(* IEC 61131-3 sources: plc-st-coding-agent/progress/evidence/f14_v10_full_20261113/jobs/custom_minimax-m27 (part 5) *)

(* ---- public-medium-05.candidate_02.st ---- *)
(* ENGINEERING_CONTRACT *)
(*
  PubRefs: PUB001, PUB003, PUB004, PUB006, PUB007
  Mode: 0=manual, 1=automatic
  Manual (Mode=FALSE): ForwardButton→MotorForward, ReverseButton→MotorReverse; interlocked (PUB001)
  Auto (Mode=TRUE):
    IDLE+SensorA→WAIT_AT_A (PUB003)
    WAIT_AT_A+ButtonA→MOVING_AB; MotorForward=TRUE (PUB003)
    MOVING_AB+SensorB→WAIT_AT_B; MotorForward=FALSE (PUB004)
    WAIT_AT_B+ButtonB→MOVING_BC; MotorForward=TRUE (PUB004)
    MOVING_BC+SensorC→WAIT_AT_C; MotorForward=FALSE (PUB004)
    WAIT_AT_C+ButtonC→COMPLETE; CompletionLight=TRUE (PUB006)
    COMPLETE+NOT SensorC→IDLE; CompletionLight=FALSE (PUB007)
  Retention: CompletionLight holds until SensorC clears (PUB007)
  Reset on mode switch: Auto state→IDLE, motor OFF
*)
(* CONTRACT_RULES [] *)

TYPE ProdState :
(
    IDLE      := 0,
    WAIT_AT_A := 1,
    MOVING_AB := 2,
    WAIT_AT_B := 3,
    MOVING_BC := 4,
    WAIT_AT_C := 5,
    COMPLETE  := 6
);
END_TYPE;

FUNCTION_BLOCK ProdLineControl
VAR_INPUT
    Mode          : BOOL;
    ForwardButton : BOOL;
    ReverseButton : BOOL;
    SensorA       : BOOL;
    SensorB       : BOOL;
    SensorC       : BOOL;
    ButtonA       : BOOL;
    ButtonB       : BOOL;
    ButtonC       : BOOL;
END_VAR
VAR
    tmp_State : ProdState := IDLE;
END_VAR
VAR_OUTPUT
    MotorForward    : BOOL := FALSE;
    MotorReverse    : BOOL := FALSE;
    CompletionLight : BOOL := FALSE;
END_VAR

// --- Automatic Mode State Machine ---
IF Mode THEN
    CASE tmp_State OF
        IDLE :
            MotorForward    := FALSE;
            MotorReverse    := FALSE;
            CompletionLight := FALSE;
            IF SensorA THEN
                tmp_State := WAIT_AT_A;
            END_IF;

        WAIT_AT_A :
            MotorForward    := FALSE;
            MotorReverse    := FALSE;
            CompletionLight := FALSE;
            IF ButtonA THEN
                tmp_State := MOVING_AB;
            END_IF;

        MOVING_AB :
            MotorForward    := TRUE;
            MotorReverse    := FALSE;
            CompletionLight := FALSE;
            IF SensorB THEN
                tmp_State     := WAIT_AT_B;
                MotorForward  := FALSE;
            END_IF;

        WAIT_AT_B :
            MotorForward    := FALSE;
            MotorReverse    := FALSE;
            CompletionLight := FALSE;
            IF ButtonB THEN
                tmp_State := MOVING_BC;
            END_IF;

        MOVING_BC :
            MotorForward    := TRUE;
            MotorReverse    := FALSE;
            CompletionLight := FALSE;
            IF SensorC THEN
                tmp_State     := WAIT_AT_C;
                MotorForward  := FALSE;
            END_IF;

        WAIT_AT_C :
            MotorForward    := FALSE;
            MotorReverse    := FALSE;
            IF ButtonC THEN
                tmp_State       := COMPLETE;
                CompletionLight := TRUE;
            END_IF;

        COMPLETE :
            MotorForward    := FALSE;
            MotorReverse    := FALSE;
            CompletionLight := TRUE;
            IF NOT SensorC THEN
                tmp_State       := IDLE;
                CompletionLight := FALSE;
            END_IF;
    END_CASE;

// --- Manual Mode ---
ELSE
    MotorForward := ForwardButton AND NOT ReverseButton;
    MotorReverse := ReverseButton AND NOT ForwardButton;
    tmp_State    := IDLE;
END_IF;

END_FUNCTION_BLOCK

(* ---- public-medium-05.raw_candidate_01.st ---- *)
(* ENGINEERING_CONTRACT *)
(*
  PubRefs: PUB001, PUB003, PUB004, PUB006, PUB007
  Mode: 0=manual, 1=automatic
  Manual (Mode=FALSE): ForwardButton→MotorForward, ReverseButton→MotorReverse; interlocked (PUB001)
  Auto (Mode=TRUE):
    IDLE+SensorA→WAIT_AT_A (PUB003)
    WAIT_AT_A+ButtonA→MOVING_AB; MotorForward=TRUE (PUB003)
    MOVING_AB+SensorB→WAIT_AT_B; MotorForward=FALSE (PUB004)
    WAIT_AT_B+ButtonB→MOVING_BC; MotorForward=TRUE (PUB004)
    MOVING_BC+SensorC→WAIT_AT_C; MotorForward=FALSE (PUB004)
    WAIT_AT_C+ButtonC→COMPLETE; CompletionLight=TRUE (PUB006)
    COMPLETE+NOT SensorC→IDLE; CompletionLight=FALSE (PUB007)
  Retention: CompletionLight holds until SensorC clears (PUB007)
  Reset on mode switch: Auto state→IDLE, motor OFF
*)
(* CONTRACT_RULES [] *)

TYPE ProdState :
(
    IDLE      := 0,
    WAIT_AT_A := 1,
    MOVING_AB := 2,
    WAIT_AT_B := 3,
    MOVING_BC := 4,
    WAIT_AT_C := 5,
    COMPLETE  := 6
);
END_TYPE

FUNCTION_BLOCK ProdLineControl
VAR
    tmp_State : ProdState := IDLE;
END_VAR
VAR_OUTPUT
    MotorForward    : BOOL := FALSE;
    MotorReverse    : BOOL := FALSE;
    CompletionLight : BOOL := FALSE;
END_VAR

// --- Automatic Mode State Machine ---
IF Mode THEN
    CASE tmp_State OF
        IDLE :
            MotorForward    := FALSE;
            MotorReverse    := FALSE;
            CompletionLight := FALSE;
            IF SensorA THEN
                tmp_State := WAIT_AT_A;
            END_IF;

        WAIT_AT_A :
            MotorForward    := FALSE;
            MotorReverse    := FALSE;
            CompletionLight := FALSE;
            IF ButtonA THEN
                tmp_State := MOVING_AB;
            END_IF;

        MOVING_AB :
            MotorForward    := TRUE;
            MotorReverse    := FALSE;
            CompletionLight := FALSE;
            IF SensorB THEN
                tmp_State     := WAIT_AT_B;
                MotorForward  := FALSE;
            END_IF;

        WAIT_AT_B :
            MotorForward    := FALSE;
            MotorReverse    := FALSE;
            CompletionLight := FALSE;
            IF ButtonB THEN
                tmp_State := MOVING_BC;
            END_IF;

        MOVING_BC :
            MotorForward    := TRUE;
            MotorReverse    := FALSE;
            CompletionLight := FALSE;
            IF SensorC THEN
                tmp_State     := WAIT_AT_C;
                MotorForward  := FALSE;
            END_IF;

        WAIT_AT_C :
            MotorForward    := FALSE;
            MotorReverse    := FALSE;
            IF ButtonC THEN
                tmp_State      := COMPLETE;
                CompletionLight := TRUE;
            END_IF;

        COMPLETE :
            MotorForward    := FALSE;
            MotorReverse    := FALSE;
            CompletionLight := TRUE;
            IF NOT SensorC THEN
                tmp_State      := IDLE;
                CompletionLight := FALSE;
            END_IF;
    END_CASE;

// --- Manual Mode ---
ELSE
    MotorForward := ForwardButton AND NOT ReverseButton;
    MotorReverse := ReverseButton AND NOT ForwardButton;
    tmp_State    := IDLE;
END_IF;

END_FUNCTION_BLOCK

(* ---- public-medium-05.raw_candidate_02.st ---- *)
(* ENGINEERING_CONTRACT *)
(*
  PubRefs: PUB001, PUB003, PUB004, PUB006, PUB007
  Mode: 0=manual, 1=automatic
  Manual (Mode=FALSE): ForwardButton→MotorForward, ReverseButton→MotorReverse; interlocked (PUB001)
  Auto (Mode=TRUE):
    IDLE+SensorA→WAIT_AT_A (PUB003)
    WAIT_AT_A+ButtonA→MOVING_AB; MotorForward=TRUE (PUB003)
    MOVING_AB+SensorB→WAIT_AT_B; MotorForward=FALSE (PUB004)
    WAIT_AT_B+ButtonB→MOVING_BC; MotorForward=TRUE (PUB004)
    MOVING_BC+SensorC→WAIT_AT_C; MotorForward=FALSE (PUB004)
    WAIT_AT_C+ButtonC→COMPLETE; CompletionLight=TRUE (PUB006)
    COMPLETE+NOT SensorC→IDLE; CompletionLight=FALSE (PUB007)
  Retention: CompletionLight holds until SensorC clears (PUB007)
  Reset on mode switch: Auto state→IDLE, motor OFF
*)
(* CONTRACT_RULES [] *)

TYPE ProdState :
(
    IDLE      := 0,
    WAIT_AT_A := 1,
    MOVING_AB := 2,
    WAIT_AT_B := 3,
    MOVING_BC := 4,
    WAIT_AT_C := 5,
    COMPLETE  := 6
);
END_TYPE;

FUNCTION_BLOCK ProdLineControl
VAR_INPUT
    Mode          : BOOL;
    ForwardButton : BOOL;
    ReverseButton : BOOL;
    SensorA       : BOOL;
    SensorB       : BOOL;
    SensorC       : BOOL;
    ButtonA       : BOOL;
    ButtonB       : BOOL;
    ButtonC       : BOOL;
END_VAR
VAR
    tmp_State : ProdState := IDLE;
END_VAR
VAR_OUTPUT
    MotorForward    : BOOL := FALSE;
    MotorReverse    : BOOL := FALSE;
    CompletionLight : BOOL := FALSE;
END_VAR

// --- Automatic Mode State Machine ---
IF Mode THEN
    CASE tmp_State OF
        IDLE :
            MotorForward    := FALSE;
            MotorReverse    := FALSE;
            CompletionLight := FALSE;
            IF SensorA THEN
                tmp_State := WAIT_AT_A;
            END_IF;

        WAIT_AT_A :
            MotorForward    := FALSE;
            MotorReverse    := FALSE;
            CompletionLight := FALSE;
            IF ButtonA THEN
                tmp_State := MOVING_AB;
            END_IF;

        MOVING_AB :
            MotorForward    := TRUE;
            MotorReverse    := FALSE;
            CompletionLight := FALSE;
            IF SensorB THEN
                tmp_State     := WAIT_AT_B;
                MotorForward  := FALSE;
            END_IF;

        WAIT_AT_B :
            MotorForward    := FALSE;
            MotorReverse    := FALSE;
            CompletionLight := FALSE;
            IF ButtonB THEN
                tmp_State := MOVING_BC;
            END_IF;

        MOVING_BC :
            MotorForward    := TRUE;
            MotorReverse    := FALSE;
            CompletionLight := FALSE;
            IF SensorC THEN
                tmp_State     := WAIT_AT_C;
                MotorForward  := FALSE;
            END_IF;

        WAIT_AT_C :
            MotorForward    := FALSE;
            MotorReverse    := FALSE;
            IF ButtonC THEN
                tmp_State       := COMPLETE;
                CompletionLight := TRUE;
            END_IF;

        COMPLETE :
            MotorForward    := FALSE;
            MotorReverse    := FALSE;
            CompletionLight := TRUE;
            IF NOT SensorC THEN
                tmp_State       := IDLE;
                CompletionLight := FALSE;
            END_IF;
    END_CASE;

// --- Manual Mode ---
ELSE
    MotorForward := ForwardButton AND NOT ReverseButton;
    MotorReverse := ReverseButton AND NOT ForwardButton;
    tmp_State    := IDLE;
END_IF;

END_FUNCTION_BLOCK

(* ---- public-medium-06.candidate_01.st ---- *)
(* ENGINEERING_CONTRACT *)
(*
| Output/State            | Activation              | Retention          | Reset/Deactivation                | Same-scan Priority | Units/Boundaries     |
|-------------------------|-------------------------|--------------------|-----------------------------------|--------------------|----------------------|
| THICKNESS_ALARM         | Immediate on valid TRUE | Hold >=500ms min   | Signal invalid OR hold timer done | Alarm active wins  | TON PT=500ms         |
| Slab_Fault_Counter      | Rising edge of valid    | Count accumulates  | Power-up only                     | N/A                | UINT max             |
| Slab_Fault_History[0]   | Rising edge of valid    | Newest entry       | Power-up only                     | N/A                | DINT timestamp       |
| Slab_Fault_History[1-4] | Shifted from lower idx  | Older entries      | Power-up only                     | N/A                | DINT timestamp       |
| Slab_Runtime_Accumulator| Accum when cutting valid| Accumulates       | Power-up only                     | N/A                | LTIME nanoseconds    |
| Hold timer (TON)        | Starts on fault clear   | Runs for PT        | Q=TRUE stops hold; signal invalid | N/A                | PT=T#500ms           |
| prev_valid_fault (VAR)  | Updated each scan       | Last cycle fault   | Power-up only                     | N/A                | BOOL                 |
| alarm_state (VAR)       | Transitions per FSM     | Holds across scans | Signal invalid resets             | N/A                | (0,1,2) enum         |
*)
(* CONTRACT_RULES [] *)

TYPE AlarmState :
(
    AlarmOff    := 0,
    FaultActive := 1,
    FaultCleared := 2
);
END_TYPE;

FUNCTION_BLOCK SlabThicknessMonitor
    VAR_INPUT
        THICKNESS_FAULT        : BOOL;
        THICKNESS_SIGNAL_VALID : BOOL;
        CUTTING_RUN            : BOOL;
        FaultTimestamp         : DINT;
        CycleTime              : TIME;
    END_VAR
    VAR_OUTPUT
        THICKNESS_ALARM         : BOOL := FALSE;
        Slab_Fault_Counter      : UINT := 0;
        Slab_Runtime_Accumulator: LTIME := LTIME#0s;
        Slab_Fault_History      : ARRAY[0..4] OF DINT := [5(DINT#0)];
    END_VAR
    VAR
        prev_valid_fault : BOOL := FALSE;
        hold_timer       : TON;
        alarm_state      : AlarmState := AlarmOff;
        tmp_hold_q       : BOOL;
    END_VAR

    // Clear all state when signal becomes invalid (power-up also covered by first-scan initialization)
    IF NOT THICKNESS_SIGNAL_VALID THEN
        alarm_state         := AlarmOff;
        THICKNESS_ALARM     := FALSE;
        hold_timer(IN := FALSE);
        prev_valid_fault    := FALSE;
        Slab_Fault_Counter  := 0;
        Slab_Fault_History  := [5(DINT#0)];
        Slab_Runtime_Accumulator := LTIME#0s;
    ELSE
        // Detect FALSE-to-TRUE transition of valid fault signal (PUB001)
        IF prev_valid_fault = FALSE AND THICKNESS_FAULT = TRUE THEN
            // Shift history: older entries toward higher indices, retain 5 most recent
            Slab_Fault_History[4] := Slab_Fault_History[3];
            Slab_Fault_History[3] := Slab_Fault_History[2];
            Slab_Fault_History[2] := Slab_Fault_History[1];
            Slab_Fault_History[1] := Slab_Fault_History[0];
            Slab_Fault_History[0] := FaultTimestamp;
            Slab_Fault_Counter := Slab_Fault_Counter + UINT#1;
        END_IF;

        // Accumulate runtime only while cutting, signal valid, no fault (PUB003)
        IF CUTTING_RUN AND NOT THICKNESS_FAULT THEN
            Slab_Runtime_Accumulator := Slab_Runtime_Accumulator + CycleTime;
        END_IF;

        // Alarm state machine with 500ms minimum hold (PUB001, PUB002)
        // Evaluate timer first so same-scan enable and elapsed origin agree
        hold_timer(IN := (alarm_state = FaultCleared));
        tmp_hold_q := hold_timer.Q;

        CASE alarm_state OF
            AlarmOff:
                IF THICKNESS_FAULT THEN
                    alarm_state     := FaultActive;
                    THICKNESS_ALARM := TRUE;
                END_IF;

            FaultActive:
                THICKNESS_ALARM := TRUE;
                IF NOT THICKNESS_FAULT THEN
                    alarm_state := FaultCleared;
                END_IF;

            FaultCleared:
                THICKNESS_ALARM := TRUE;
                IF tmp_hold_q THEN
                    alarm_state     := AlarmOff;
                    THICKNESS_ALARM := FALSE;
                END_IF;
        END_CASE;
    END_IF;

    // Update previous fault state for next scan edge detection
    prev_valid_fault := THICKNESS_FAULT;
END_FUNCTION_BLOCK

(* ---- public-medium-06.candidate_02.st ---- *)
(* ENGINEERING_CONTRACT *)
(*
| Output/State            | Activation              | Retention          | Reset/Deactivation                | Same-scan Priority | Units/Boundaries     |
|-------------------------|-------------------------|--------------------|-----------------------------------|--------------------|----------------------|
| THICKNESS_ALARM         | Immediate on valid TRUE | Hold >=500ms min   | Signal invalid OR hold timer done | Alarm active wins  | TON PT=500ms         |
| Slab_Fault_Counter      | Rising edge of valid    | Count accumulates  | Power-up only                     | N/A                | UINT max             |
| Slab_Fault_History[0]   | Rising edge of valid    | Newest entry       | Power-up only                     | N/A                | DINT timestamp       |
| Slab_Fault_History[1-4] | Shifted from lower idx  | Older entries      | Power-up only                     | N/A                | DINT timestamp       |
| Slab_Runtime_Accumulator| Accum when cutting valid| Accumulates       | Power-up only                     | N/A                | LTIME nanoseconds    |
| Hold timer (TON)        | Starts on fault clear   | Runs for PT        | Q=TRUE stops hold; signal invalid | N/A                | PT=T#500ms           |
| prev_valid_fault (VAR)  | Updated each scan       | Last cycle fault   | Power-up only                     | N/A                | BOOL                 |
| alarm_state (VAR)       | Transitions per FSM     | Holds across scans | Signal invalid resets             | N/A                | (0,1,2) enum         |
*)
(* CONTRACT_RULES [] *)

TYPE AlarmState :
(
    AlarmOff    := 0,
    FaultActive := 1,
    FaultCleared := 2
);
END_TYPE;

FUNCTION_BLOCK SlabThicknessMonitor
    VAR_INPUT
        THICKNESS_FAULT        : BOOL;
        THICKNESS_SIGNAL_VALID : BOOL;
        CUTTING_RUN            : BOOL;
        FaultTimestamp         : DINT;
        CycleTime              : TIME;
    END_VAR
    VAR_OUTPUT
        THICKNESS_ALARM         : BOOL := FALSE;
        Slab_Fault_Counter      : UINT := 0;
        Slab_Runtime_Accumulator: LTIME := LTIME#0s;
        Slab_Fault_History      : ARRAY[0..4] OF DINT := [DINT#0, DINT#0, DINT#0, DINT#0, DINT#0];
    END_VAR
    VAR
        prev_valid_fault : BOOL := FALSE;
        hold_timer       : TON;
        alarm_state      : AlarmState := AlarmOff;
        tmp_hold_q       : BOOL;
    END_VAR

    // Clear all state when signal becomes invalid (power-up also covered by first-scan initialization)
    IF NOT THICKNESS_SIGNAL_VALID THEN
        alarm_state         := AlarmOff;
        THICKNESS_ALARM     := FALSE;
        hold_timer(IN := FALSE);
        prev_valid_fault    := FALSE;
        Slab_Fault_Counter  := 0;
        Slab_Fault_History  := [DINT#0, DINT#0, DINT#0, DINT#0, DINT#0];
        Slab_Runtime_Accumulator := LTIME#0s;
    ELSE
        // Detect FALSE-to-TRUE transition of valid fault signal (PUB001)
        IF prev_valid_fault = FALSE AND THICKNESS_FAULT = TRUE THEN
            // Shift history: older entries toward higher indices, retain 5 most recent
            Slab_Fault_History[4] := Slab_Fault_History[3];
            Slab_Fault_History[3] := Slab_Fault_History[2];
            Slab_Fault_History[2] := Slab_Fault_History[1];
            Slab_Fault_History[1] := Slab_Fault_History[0];
            Slab_Fault_History[0] := FaultTimestamp;
            Slab_Fault_Counter := Slab_Fault_Counter + UINT#1;
        END_IF;

        // Accumulate runtime only while cutting, signal valid, no fault (PUB003)
        IF CUTTING_RUN AND NOT THICKNESS_FAULT THEN
            Slab_Runtime_Accumulator := Slab_Runtime_Accumulator + CycleTime;
        END_IF;

        // Alarm state machine with 500ms minimum hold (PUB001, PUB002)
        // Evaluate timer first so same-scan enable and elapsed origin agree
        hold_timer(IN := (alarm_state = FaultCleared));
        tmp_hold_q := hold_timer.Q;

        CASE alarm_state OF
            AlarmOff:
                IF THICKNESS_FAULT THEN
                    alarm_state     := FaultActive;
                    THICKNESS_ALARM := TRUE;
                END_IF;

            FaultActive:
                THICKNESS_ALARM := TRUE;
                IF NOT THICKNESS_FAULT THEN
                    alarm_state := FaultCleared;
                END_IF;

            FaultCleared:
                THICKNESS_ALARM := TRUE;
                IF tmp_hold_q THEN
                    alarm_state     := AlarmOff;
                    THICKNESS_ALARM := FALSE;
                END_IF;
        END_CASE;
    END_IF;

    // Update previous fault state for next scan edge detection
    prev_valid_fault := THICKNESS_FAULT;
END_FUNCTION_BLOCK

(* ---- public-medium-06.candidate_03.st ---- *)
(* ENGINEERING_CONTRACT *)
(*
| Output/State            | Activation              | Retention          | Reset/Deactivation                | Same-scan Priority | Units/Boundaries     |
|-------------------------|-------------------------|--------------------|-----------------------------------|--------------------|----------------------|
| THICKNESS_ALARM         | Immediate on valid TRUE | Hold >=500ms min   | Signal invalid OR hold timer done | Alarm active wins  | TON PT=500ms         |
| Slab_Fault_Counter      | Rising edge of valid    | Count accumulates  | Power-up only                     | N/A                | UINT max             |
| Slab_Fault_History[0]   | Rising edge of valid    | Newest entry       | Power-up only                     | N/A                | DINT timestamp       |
| Slab_Fault_History[1-4] | Shifted from lower idx  | Older entries      | Power-up only                     | N/A                | DINT timestamp       |
| Slab_Runtime_Accumulator| Accum when cutting valid| Accumulates       | Power-up only                     | N/A                | LTIME nanoseconds    |
| Hold timer (TON)        | Starts on fault clear   | Runs for PT        | Q=TRUE stops hold; signal invalid | N/A                | PT=T#500ms           |
| prev_valid_fault (VAR)  | Updated each scan       | Last cycle fault   | Power-up only                     | N/A                | BOOL                 |
| alarm_state (VAR)       | Transitions per FSM     | Holds across scans | Signal invalid resets             | N/A                | (0,1,2) enum         |
*)
(* CONTRACT_RULES [] *)

TYPE AlarmState :
(
    AlarmOff    := 0,
    FaultActive := 1,
    FaultCleared := 2
);
END_TYPE;

FUNCTION_BLOCK SlabThicknessMonitor
    VAR_INPUT
        THICKNESS_FAULT        : BOOL;
        THICKNESS_SIGNAL_VALID : BOOL;
        CUTTING_RUN            : BOOL;
        FaultTimestamp         : DINT;
        CycleTime              : TIME;
    END_VAR
    VAR_OUTPUT
        THICKNESS_ALARM         : BOOL := FALSE;
        Slab_Fault_Counter      : UINT := 0;
        Slab_Runtime_Accumulator: LTIME := LTIME#0s;
        Slab_Fault_History      : ARRAY[0..4] OF DINT;
    END_VAR
    VAR
        prev_valid_fault : BOOL := FALSE;
        hold_timer       : TON;
        alarm_state      : AlarmState := AlarmOff;
        tmp_hold_q       : BOOL;
        tmp_idx          : UINT;
    END_VAR

    // Clear all state when signal becomes invalid (power-up also covered by first-scan initialization)
    IF NOT THICKNESS_SIGNAL_VALID THEN
        alarm_state         := AlarmOff;
        THICKNESS_ALARM     := FALSE;
        hold_timer(IN := FALSE);
        prev_valid_fault    := FALSE;
        Slab_Fault_Counter  := 0;
        Slab_Fault_History[0] := DINT#0;
        Slab_Fault_History[1] := DINT#0;
        Slab_Fault_History[2] := DINT#0;
        Slab_Fault_History[3] := DINT#0;
        Slab_Fault_History[4] := DINT#0;
        Slab_Runtime_Accumulator := LTIME#0s;
    ELSE
        // Detect FALSE-to-TRUE transition of valid fault signal (PUB001)
        IF prev_valid_fault = FALSE AND THICKNESS_FAULT = TRUE THEN
            // Shift history: older entries toward higher indices, retain 5 most recent
            Slab_Fault_History[4] := Slab_Fault_History[3];
            Slab_Fault_History[3] := Slab_Fault_History[2];
            Slab_Fault_History[2] := Slab_Fault_History[1];
            Slab_Fault_History[1] := Slab_Fault_History[0];
            Slab_Fault_History[0] := FaultTimestamp;
            Slab_Fault_Counter := Slab_Fault_Counter + UINT#1;
        END_IF;

        // Accumulate runtime only while cutting, signal valid, no fault (PUB003)
        IF CUTTING_RUN AND NOT THICKNESS_FAULT THEN
            Slab_Runtime_Accumulator := Slab_Runtime_Accumulator + CycleTime;
        END_IF;

        // Alarm state machine with 500ms minimum hold (PUB001, PUB002)
        // Evaluate timer first so same-scan enable and elapsed origin agree
        hold_timer(IN := (alarm_state = FaultCleared));
        tmp_hold_q := hold_timer.Q;

        CASE alarm_state OF
            AlarmOff:
                IF THICKNESS_FAULT THEN
                    alarm_state     := FaultActive;
                    THICKNESS_ALARM := TRUE;
                END_IF;

            FaultActive:
                THICKNESS_ALARM := TRUE;
                IF NOT THICKNESS_FAULT THEN
                    alarm_state := FaultCleared;
                END_IF;

            FaultCleared:
                THICKNESS_ALARM := TRUE;
                IF tmp_hold_q THEN
                    alarm_state     := AlarmOff;
                    THICKNESS_ALARM := FALSE;
                END_IF;
        END_CASE;
    END_IF;

    // Update previous fault state for next scan edge detection
    prev_valid_fault := THICKNESS_FAULT;
END_FUNCTION_BLOCK

(* ---- public-medium-06.candidate_04.st ---- *)
(* ENGINEERING_CONTRACT *)
(*
| Output/State            | Activation              | Retention          | Reset/Deactivation                | Same-scan Priority | Units/Boundaries     |
|-------------------------|-------------------------|--------------------|-----------------------------------|--------------------|----------------------|
| THICKNESS_ALARM         | Immediate on valid TRUE | Hold >=500ms min   | Signal invalid OR hold timer done | Alarm active wins  | TON PT=T#500ms       |
| Slab_Fault_Counter      | Rising edge of valid    | Count accumulates  | Power-up only                     | N/A                | UINT max             |
| Slab_Fault_History[0]   | Rising edge of valid    | Newest entry       | Power-up only                     | N/A                | DINT timestamp       |
| Slab_Fault_History[1-4] | Shifted from lower idx  | Older entries      | Power-up only                     | N/A                | DINT timestamp       |
| Slab_Runtime_Accumulator| Accum when cutting valid| Accumulates       | Power-up only                     | N/A                | LTIME nanoseconds    |
| Hold timer (TON)        | Starts on fault clear   | Runs for PT        | Q=TRUE stops hold; signal invalid | N/A                | PT=T#500ms           |
| prev_valid_fault (VAR)  | Updated each scan       | Last cycle fault   | Power-up only                     | N/A                | BOOL                 |
| alarm_state (VAR)       | Transitions per FSM     | Holds across scans | Signal invalid resets             | N/A                | (0,1,2) enum         |
*)
(* CONTRACT_RULES [] *)

TYPE AlarmState :
(
    AlarmOff    := 0,
    FaultActive := 1,
    FaultCleared := 2
);
END_TYPE;

FUNCTION_BLOCK SlabThicknessMonitor
    VAR_INPUT
        THICKNESS_FAULT        : BOOL;
        THICKNESS_SIGNAL_VALID : BOOL;
        CUTTING_RUN            : BOOL;
        FaultTimestamp         : DINT;
        CycleTime              : TIME;
    END_VAR
    VAR_OUTPUT
        THICKNESS_ALARM         : BOOL := FALSE;
        Slab_Fault_Counter      : UINT := 0;
        Slab_Runtime_Accumulator: LTIME := LTIME#0s;
        Slab_Fault_History      : ARRAY[0..4] OF DINT;
    END_VAR
    VAR
        prev_valid_fault : BOOL := FALSE;
        hold_timer       : TON;
        alarm_state      : AlarmState := AlarmOff;
        tmp_hold_q       : BOOL;
        tmp_idx          : UINT;
    END_VAR

    // Clear all state when signal becomes invalid (power-up also covered by first-scan initialization)
    IF NOT THICKNESS_SIGNAL_VALID THEN
        alarm_state         := AlarmOff;
        THICKNESS_ALARM     := FALSE;
        prev_valid_fault    := FALSE;
        Slab_Fault_Counter  := 0;
        Slab_Fault_History[0] := DINT#0;
        Slab_Fault_History[1] := DINT#0;
        Slab_Fault_History[2] := DINT#0;
        Slab_Fault_History[3] := DINT#0;
        Slab_Fault_History[4] := DINT#0;
        Slab_Runtime_Accumulator := LTIME#0s;
        hold_timer(IN := FALSE, PT := T#500ms, RESET := TRUE);
    ELSE
        // Detect FALSE-to-TRUE transition of valid fault signal (PUB001)
        IF prev_valid_fault = FALSE AND THICKNESS_FAULT = TRUE THEN
            // Shift history: older entries toward higher indices, retain 5 most recent
            Slab_Fault_History[4] := Slab_Fault_History[3];
            Slab_Fault_History[3] := Slab_Fault_History[2];
            Slab_Fault_History[2] := Slab_Fault_History[1];
            Slab_Fault_History[1] := Slab_Fault_History[0];
            Slab_Fault_History[0] := FaultTimestamp;
            Slab_Fault_Counter := Slab_Fault_Counter + UINT#1;
        END_IF;

        // Accumulate runtime only while cutting, signal valid, no fault (PUB003)
        IF CUTTING_RUN AND NOT THICKNESS_FAULT THEN
            Slab_Runtime_Accumulator := Slab_Runtime_Accumulator + TIME_TO_LTIME(CycleTime);
        END_IF;

        // Alarm state machine with 500ms minimum hold (PUB001, PUB002)
        // Evaluate timer first so same-scan enable and elapsed origin agree
        hold_timer(IN := (alarm_state = FaultCleared), PT := T#500ms, RESET := FALSE);
        tmp_hold_q := hold_timer.Q;

        CASE alarm_state OF
            AlarmOff:
                IF THICKNESS_FAULT THEN
                    alarm_state     := FaultActive;
                    THICKNESS_ALARM := TRUE;
                END_IF;

            FaultActive:
                THICKNESS_ALARM := TRUE;
                IF NOT THICKNESS_FAULT THEN
                    alarm_state := FaultCleared;
                END_IF;

            FaultCleared:
                THICKNESS_ALARM := TRUE;
                IF tmp_hold_q THEN
                    alarm_state     := AlarmOff;
                    THICKNESS_ALARM := FALSE;
                END_IF;
        END_CASE;
    END_IF;

    // Update previous fault state for next scan edge detection
    prev_valid_fault := THICKNESS_FAULT;
END_FUNCTION_BLOCK

(* ---- public-medium-06.raw_candidate_01.st ---- *)
(* ENGINEERING_CONTRACT *)
(*
| Output/State            | Activation              | Retention          | Reset/Deactivation                | Same-scan Priority | Units/Boundaries     |
|-------------------------|-------------------------|--------------------|-----------------------------------|--------------------|----------------------|
| THICKNESS_ALARM         | Immediate on valid TRUE | Hold >=500ms min   | Signal invalid OR hold timer done | Alarm active wins  | TON PT=500ms         |
| Slab_Fault_Counter      | Rising edge of valid    | Count accumulates  | Power-up only                     | N/A                | UINT max             |
| Slab_Fault_History[0]   | Rising edge of valid    | Newest entry       | Power-up only                     | N/A                | DINT timestamp       |
| Slab_Fault_History[1-4] | Shifted from lower idx  | Older entries      | Power-up only                     | N/A                | DINT timestamp       |
| Slab_Runtime_Accumulator| Accum when cutting valid| Accumulates       | Power-up only                     | N/A                | LTIME nanoseconds    |
| Hold timer (TON)        | Starts on fault clear   | Runs for PT        | Q=TRUE stops hold; signal invalid | N/A                | PT=T#500ms           |
| prev_valid_fault (VAR)  | Updated each scan       | Last cycle fault   | Power-up only                     | N/A                | BOOL                 |
| alarm_state (VAR)       | Transitions per FSM     | Holds across scans | Signal invalid resets             | N/A                | (0,1,2) enum         |
*)
(* CONTRACT_RULES [] *)

TYPE AlarmState :
(
    AlarmOff    := 0,
    FaultActive := 1,
    FaultCleared := 2
);
END_TYPE

FUNCTION_BLOCK SlabThicknessMonitor
    VAR_INPUT
        THICKNESS_FAULT        : BOOL;
        THICKNESS_SIGNAL_VALID : BOOL;
        CUTTING_RUN            : BOOL;
        FaultTimestamp         : DINT;
        CycleTime              : TIME;
    END_VAR
    VAR_OUTPUT
        THICKNESS_ALARM         : BOOL := FALSE;
        Slab_Fault_Counter      : UINT := 0;
        Slab_Runtime_Accumulator: LTIME := LTIME#0s;
        Slab_Fault_History      : ARRAY[0..4] OF DINT := [5(DINT#0)];
    END_VAR
    VAR
        prev_valid_fault : BOOL := FALSE;
        hold_timer       : TON;
        alarm_state      : AlarmState := AlarmOff;
        tmp_hold_q       : BOOL;
    END_VAR

    // Clear all state when signal becomes invalid (power-up also covered by first-scan initialization)
    IF NOT THICKNESS_SIGNAL_VALID THEN
        alarm_state         := AlarmOff;
        THICKNESS_ALARM     := FALSE;
        hold_timer(IN := FALSE);
        prev_valid_fault    := FALSE;
        Slab_Fault_Counter  := 0;
        Slab_Fault_History  := [5(DINT#0)];
        Slab_Runtime_Accumulator := LTIME#0s;
    ELSE
        // Detect FALSE-to-TRUE transition of valid fault signal (PUB001)
        IF prev_valid_fault = FALSE AND THICKNESS_FAULT = TRUE THEN
            // Shift history: older entries toward higher indices, retain 5 most recent
            Slab_Fault_History[4] := Slab_Fault_History[3];
            Slab_Fault_History[3] := Slab_Fault_History[2];
            Slab_Fault_History[2] := Slab_Fault_History[1];
            Slab_Fault_History[1] := Slab_Fault_History[0];
            Slab_Fault_History[0] := FaultTimestamp;
            Slab_Fault_Counter := Slab_Fault_Counter + UINT#1;
        END_IF

        // Accumulate runtime only while cutting, signal valid, no fault (PUB003)
        IF CUTTING_RUN AND NOT THICKNESS_FAULT THEN
            Slab_Runtime_Accumulator := Slab_Runtime_Accumulator + CycleTime;
        END_IF

        // Alarm state machine with 500ms minimum hold (PUB001, PUB002)
        // Evaluate timer first so same-scan enable and elapsed origin agree
        hold_timer(IN := (alarm_state = FaultCleared));
        tmp_hold_q := hold_timer.Q;

        CASE alarm_state OF
            AlarmOff:
                IF THICKNESS_FAULT THEN
                    alarm_state     := FaultActive;
                    THICKNESS_ALARM := TRUE;
                END_IF;

            FaultActive:
                THICKNESS_ALARM := TRUE;
                IF NOT THICKNESS_FAULT THEN
                    alarm_state := FaultCleared;
                END_IF;

            FaultCleared:
                THICKNESS_ALARM := TRUE;
                IF tmp_hold_q THEN
                    alarm_state     := AlarmOff;
                    THICKNESS_ALARM := FALSE;
                END_IF;
        END_CASE;
    END_IF;

    // Update previous fault state for next scan edge detection
    prev_valid_fault := THICKNESS_FAULT;
END_FUNCTION_BLOCK

(* ---- public-medium-06.raw_candidate_02.st ---- *)
(* ENGINEERING_CONTRACT *)
(*
| Output/State            | Activation              | Retention          | Reset/Deactivation                | Same-scan Priority | Units/Boundaries     |
|-------------------------|-------------------------|--------------------|-----------------------------------|--------------------|----------------------|
| THICKNESS_ALARM         | Immediate on valid TRUE | Hold >=500ms min   | Signal invalid OR hold timer done | Alarm active wins  | TON PT=500ms         |
| Slab_Fault_Counter      | Rising edge of valid    | Count accumulates  | Power-up only                     | N/A                | UINT max             |
| Slab_Fault_History[0]   | Rising edge of valid    | Newest entry       | Power-up only                     | N/A                | DINT timestamp       |
| Slab_Fault_History[1-4] | Shifted from lower idx  | Older entries      | Power-up only                     | N/A                | DINT timestamp       |
| Slab_Runtime_Accumulator| Accum when cutting valid| Accumulates       | Power-up only                     | N/A                | LTIME nanoseconds    |
| Hold timer (TON)        | Starts on fault clear   | Runs for PT        | Q=TRUE stops hold; signal invalid | N/A                | PT=T#500ms           |
| prev_valid_fault (VAR)  | Updated each scan       | Last cycle fault   | Power-up only                     | N/A                | BOOL                 |
| alarm_state (VAR)       | Transitions per FSM     | Holds across scans | Signal invalid resets             | N/A                | (0,1,2) enum         |
*)
(* CONTRACT_RULES [] *)

TYPE AlarmState :
(
    AlarmOff    := 0,
    FaultActive := 1,
    FaultCleared := 2
);
END_TYPE;

FUNCTION_BLOCK SlabThicknessMonitor
    VAR_INPUT
        THICKNESS_FAULT        : BOOL;
        THICKNESS_SIGNAL_VALID : BOOL;
        CUTTING_RUN            : BOOL;
        FaultTimestamp         : DINT;
        CycleTime              : TIME;
    END_VAR
    VAR_OUTPUT
        THICKNESS_ALARM         : BOOL := FALSE;
        Slab_Fault_Counter      : UINT := 0;
        Slab_Runtime_Accumulator: LTIME := LTIME#0s;
        Slab_Fault_History      : ARRAY[0..4] OF DINT := [DINT#0, DINT#0, DINT#0, DINT#0, DINT#0];
    END_VAR
    VAR
        prev_valid_fault : BOOL := FALSE;
        hold_timer       : TON;
        alarm_state      : AlarmState := AlarmOff;
        tmp_hold_q       : BOOL;
    END_VAR

    // Clear all state when signal becomes invalid (power-up also covered by first-scan initialization)
    IF NOT THICKNESS_SIGNAL_VALID THEN
        alarm_state         := AlarmOff;
        THICKNESS_ALARM     := FALSE;
        hold_timer(IN := FALSE);
        prev_valid_fault    := FALSE;
        Slab_Fault_Counter  := 0;
        Slab_Fault_History  := [DINT#0, DINT#0, DINT#0, DINT#0, DINT#0];
        Slab_Runtime_Accumulator := LTIME#0s;
    ELSE
        // Detect FALSE-to-TRUE transition of valid fault signal (PUB001)
        IF prev_valid_fault = FALSE AND THICKNESS_FAULT = TRUE THEN
            // Shift history: older entries toward higher indices, retain 5 most recent
            Slab_Fault_History[4] := Slab_Fault_History[3];
            Slab_Fault_History[3] := Slab_Fault_History[2];
            Slab_Fault_History[2] := Slab_Fault_History[1];
            Slab_Fault_History[1] := Slab_Fault_History[0];
            Slab_Fault_History[0] := FaultTimestamp;
            Slab_Fault_Counter := Slab_Fault_Counter + UINT#1;
        END_IF;

        // Accumulate runtime only while cutting, signal valid, no fault (PUB003)
        IF CUTTING_RUN AND NOT THICKNESS_FAULT THEN
            Slab_Runtime_Accumulator := Slab_Runtime_Accumulator + CycleTime;
        END_IF;

        // Alarm state machine with 500ms minimum hold (PUB001, PUB002)
        // Evaluate timer first so same-scan enable and elapsed origin agree
        hold_timer(IN := (alarm_state = FaultCleared));
        tmp_hold_q := hold_timer.Q;

        CASE alarm_state OF
            AlarmOff:
                IF THICKNESS_FAULT THEN
                    alarm_state     := FaultActive;
                    THICKNESS_ALARM := TRUE;
                END_IF;

            FaultActive:
                THICKNESS_ALARM := TRUE;
                IF NOT THICKNESS_FAULT THEN
                    alarm_state := FaultCleared;
                END_IF;

            FaultCleared:
                THICKNESS_ALARM := TRUE;
                IF tmp_hold_q THEN
                    alarm_state     := AlarmOff;
                    THICKNESS_ALARM := FALSE;
                END_IF;
        END_CASE;
    END_IF;

    // Update previous fault state for next scan edge detection
    prev_valid_fault := THICKNESS_FAULT;
END_FUNCTION_BLOCK

(* ---- public-medium-06.raw_candidate_03.st ---- *)
(* ENGINEERING_CONTRACT *)
(*
| Output/State            | Activation              | Retention          | Reset/Deactivation                | Same-scan Priority | Units/Boundaries     |
|-------------------------|-------------------------|--------------------|-----------------------------------|--------------------|----------------------|
| THICKNESS_ALARM         | Immediate on valid TRUE | Hold >=500ms min   | Signal invalid OR hold timer done | Alarm active wins  | TON PT=500ms         |
| Slab_Fault_Counter      | Rising edge of valid    | Count accumulates  | Power-up only                     | N/A                | UINT max             |
| Slab_Fault_History[0]   | Rising edge of valid    | Newest entry       | Power-up only                     | N/A                | DINT timestamp       |
| Slab_Fault_History[1-4] | Shifted from lower idx  | Older entries      | Power-up only                     | N/A                | DINT timestamp       |
| Slab_Runtime_Accumulator| Accum when cutting valid| Accumulates       | Power-up only                     | N/A                | LTIME nanoseconds    |
| Hold timer (TON)        | Starts on fault clear   | Runs for PT        | Q=TRUE stops hold; signal invalid | N/A                | PT=T#500ms           |
| prev_valid_fault (VAR)  | Updated each scan       | Last cycle fault   | Power-up only                     | N/A                | BOOL                 |
| alarm_state (VAR)       | Transitions per FSM     | Holds across scans | Signal invalid resets             | N/A                | (0,1,2) enum         |
*)
(* CONTRACT_RULES [] *)

TYPE AlarmState :
(
    AlarmOff    := 0,
    FaultActive := 1,
    FaultCleared := 2
);
END_TYPE;

FUNCTION_BLOCK SlabThicknessMonitor
    VAR_INPUT
        THICKNESS_FAULT        : BOOL;
        THICKNESS_SIGNAL_VALID : BOOL;
        CUTTING_RUN            : BOOL;
        FaultTimestamp         : DINT;
        CycleTime              : TIME;
    END_VAR
    VAR_OUTPUT
        THICKNESS_ALARM         : BOOL := FALSE;
        Slab_Fault_Counter      : UINT := 0;
        Slab_Runtime_Accumulator: LTIME := LTIME#0s;
        Slab_Fault_History      : ARRAY[0..4] OF DINT;
    END_VAR
    VAR
        prev_valid_fault : BOOL := FALSE;
        hold_timer       : TON;
        alarm_state      : AlarmState := AlarmOff;
        tmp_hold_q       : BOOL;
        tmp_idx          : UINT;
    END_VAR

    // Clear all state when signal becomes invalid (power-up also covered by first-scan initialization)
    IF NOT THICKNESS_SIGNAL_VALID THEN
        alarm_state         := AlarmOff;
        THICKNESS_ALARM     := FALSE;
        hold_timer(IN := FALSE);
        prev_valid_fault    := FALSE;
        Slab_Fault_Counter  := 0;
        Slab_Fault_History[0] := DINT#0;
        Slab_Fault_History[1] := DINT#0;
        Slab_Fault_History[2] := DINT#0;
        Slab_Fault_History[3] := DINT#0;
        Slab_Fault_History[4] := DINT#0;
        Slab_Runtime_Accumulator := LTIME#0s;
    ELSE
        // Detect FALSE-to-TRUE transition of valid fault signal (PUB001)
        IF prev_valid_fault = FALSE AND THICKNESS_FAULT = TRUE THEN
            // Shift history: older entries toward higher indices, retain 5 most recent
            Slab_Fault_History[4] := Slab_Fault_History[3];
            Slab_Fault_History[3] := Slab_Fault_History[2];
            Slab_Fault_History[2] := Slab_Fault_History[1];
            Slab_Fault_History[1] := Slab_Fault_History[0];
            Slab_Fault_History[0] := FaultTimestamp;
            Slab_Fault_Counter := Slab_Fault_Counter + UINT#1;
        END_IF;

        // Accumulate runtime only while cutting, signal valid, no fault (PUB003)
        IF CUTTING_RUN AND NOT THICKNESS_FAULT THEN
            Slab_Runtime_Accumulator := Slab_Runtime_Accumulator + CycleTime;
        END_IF;

        // Alarm state machine with 500ms minimum hold (PUB001, PUB002)
        // Evaluate timer first so same-scan enable and elapsed origin agree
        hold_timer(IN := (alarm_state = FaultCleared));
        tmp_hold_q := hold_timer.Q;

        CASE alarm_state OF
            AlarmOff:
                IF THICKNESS_FAULT THEN
                    alarm_state     := FaultActive;
                    THICKNESS_ALARM := TRUE;
                END_IF;

            FaultActive:
                THICKNESS_ALARM := TRUE;
                IF NOT THICKNESS_FAULT THEN
                    alarm_state := FaultCleared;
                END_IF;

            FaultCleared:
                THICKNESS_ALARM := TRUE;
                IF tmp_hold_q THEN
                    alarm_state     := AlarmOff;
                    THICKNESS_ALARM := FALSE;
                END_IF;
        END_CASE;
    END_IF;

    // Update previous fault state for next scan edge detection
    prev_valid_fault := THICKNESS_FAULT;
END_FUNCTION_BLOCK

(* ---- public-medium-06.raw_candidate_04.st ---- *)
(* ENGINEERING_CONTRACT *)
(*
| Output/State            | Activation              | Retention          | Reset/Deactivation                | Same-scan Priority | Units/Boundaries     |
|-------------------------|-------------------------|--------------------|-----------------------------------|--------------------|----------------------|
| THICKNESS_ALARM         | Immediate on valid TRUE | Hold >=500ms min   | Signal invalid OR hold timer done | Alarm active wins  | TON PT=T#500ms       |
| Slab_Fault_Counter      | Rising edge of valid    | Count accumulates  | Power-up only                     | N/A                | UINT max             |
| Slab_Fault_History[0]   | Rising edge of valid    | Newest entry       | Power-up only                     | N/A                | DINT timestamp       |
| Slab_Fault_History[1-4] | Shifted from lower idx  | Older entries      | Power-up only                     | N/A                | DINT timestamp       |
| Slab_Runtime_Accumulator| Accum when cutting valid| Accumulates       | Power-up only                     | N/A                | LTIME nanoseconds    |
| Hold timer (TON)        | Starts on fault clear   | Runs for PT        | Q=TRUE stops hold; signal invalid | N/A                | PT=T#500ms           |
| prev_valid_fault (VAR)  | Updated each scan       | Last cycle fault   | Power-up only                     | N/A                | BOOL                 |
| alarm_state (VAR)       | Transitions per FSM     | Holds across scans | Signal invalid resets             | N/A                | (0,1,2) enum         |
*)
(* CONTRACT_RULES [] *)

TYPE AlarmState :
(
    AlarmOff    := 0,
    FaultActive := 1,
    FaultCleared := 2
);
END_TYPE;

FUNCTION_BLOCK SlabThicknessMonitor
    VAR_INPUT
        THICKNESS_FAULT        : BOOL;
        THICKNESS_SIGNAL_VALID : BOOL;
        CUTTING_RUN            : BOOL;
        FaultTimestamp         : DINT;
        CycleTime              : TIME;
    END_VAR
    VAR_OUTPUT
        THICKNESS_ALARM         : BOOL := FALSE;
        Slab_Fault_Counter      : UINT := 0;
        Slab_Runtime_Accumulator: LTIME := LTIME#0s;
        Slab_Fault_History      : ARRAY[0..4] OF DINT;
    END_VAR
    VAR
        prev_valid_fault : BOOL := FALSE;
        hold_timer       : TON;
        alarm_state      : AlarmState := AlarmOff;
        tmp_hold_q       : BOOL;
        tmp_idx          : UINT;
    END_VAR

    // Clear all state when signal becomes invalid (power-up also covered by first-scan initialization)
    IF NOT THICKNESS_SIGNAL_VALID THEN
        alarm_state         := AlarmOff;
        THICKNESS_ALARM     := FALSE;
        prev_valid_fault    := FALSE;
        Slab_Fault_Counter  := 0;
        Slab_Fault_History[0] := DINT#0;
        Slab_Fault_History[1] := DINT#0;
        Slab_Fault_History[2] := DINT#0;
        Slab_Fault_History[3] := DINT#0;
        Slab_Fault_History[4] := DINT#0;
        Slab_Runtime_Accumulator := LTIME#0s;
        hold_timer(IN := FALSE, PT := T#500ms, RESET := TRUE);
    ELSE
        // Detect FALSE-to-TRUE transition of valid fault signal (PUB001)
        IF prev_valid_fault = FALSE AND THICKNESS_FAULT = TRUE THEN
            // Shift history: older entries toward higher indices, retain 5 most recent
            Slab_Fault_History[4] := Slab_Fault_History[3];
            Slab_Fault_History[3] := Slab_Fault_History[2];
            Slab_Fault_History[2] := Slab_Fault_History[1];
            Slab_Fault_History[1] := Slab_Fault_History[0];
            Slab_Fault_History[0] := FaultTimestamp;
            Slab_Fault_Counter := Slab_Fault_Counter + UINT#1;
        END_IF;

        // Accumulate runtime only while cutting, signal valid, no fault (PUB003)
        IF CUTTING_RUN AND NOT THICKNESS_FAULT THEN
            Slab_Runtime_Accumulator := Slab_Runtime_Accumulator + TIME_TO_LTIME(CycleTime);
        END_IF;

        // Alarm state machine with 500ms minimum hold (PUB001, PUB002)
        // Evaluate timer first so same-scan enable and elapsed origin agree
        hold_timer(IN := (alarm_state = FaultCleared), PT := T#500ms, RESET := FALSE);
        tmp_hold_q := hold_timer.Q;

        CASE alarm_state OF
            AlarmOff:
                IF THICKNESS_FAULT THEN
                    alarm_state     := FaultActive;
                    THICKNESS_ALARM := TRUE;
                END_IF;

            FaultActive:
                THICKNESS_ALARM := TRUE;
                IF NOT THICKNESS_FAULT THEN
                    alarm_state := FaultCleared;
                END_IF;

            FaultCleared:
                THICKNESS_ALARM := TRUE;
                IF tmp_hold_q THEN
                    alarm_state     := AlarmOff;
                    THICKNESS_ALARM := FALSE;
                END_IF;
        END_CASE;
    END_IF;

    // Update previous fault state for next scan edge detection
    prev_valid_fault := THICKNESS_FAULT;
END_FUNCTION_BLOCK

(* ---- public-medium-07.candidate_01.st ---- *)
(* ENGINEERING_CONTRACT
 * | Output/State Group | Activation              | Retention         | Reset/Deactivation                  | Priority | Units/Bounds          |
 * |---------------------|-------------------------|-------------------|-------------------------------------|----------|-----------------------|
 * | SUPPLY_FAN_RUN      | 30s TON.Q after         | Hold TRUE while   | Deactivate and reset TON when:      | Same-scan| 30s PT, BOOLEAN       |
 * |   - Fan Start       |   Occupied=TRUE AND     |   conditions      |   Occupied=FALSE OR Mode=3 (Night)  |          |                       |
 * |                     |   Mode<>3, rising edge  |   maintained      |   Rising-edge reset on recovery     |          |                       |
 * |---------------------|-------------------------|-------------------|-------------------------------------|----------|-----------------------|
 * | TEMP_SETPOINT_ADJUST| Computed each scan from | Computed fresh    | Recalculated on any input change    | Same-scan| Auto: 0/+3/+2,        |
 * |   - Auto (Mode=0)   |   Mode × Occupancy ×    |   each scan       |   No explicit retention             |          |   Comfort: 0/+1,      |
 * |   - Comfort (Mode=1)|   EnergySaving combo    |                   |                                     |          |   Economy: 0/+4,      |
 * |   - Economy (Mode=2)|                         |                   |                                     |          |   Night: +4, ±4°C     |
 * |   - Night (Mode=3)  |                         |                   |                                     |          |                       |
 * PUB clause citations: PUB001, PUB002, PUB003, PUB004, PUB005, PUB006, PUB007, PUB008
 *)

(* CONTRACT_RULES [] *)

FUNCTION_BLOCK FB_HVAC_Control
VAR
    local_TON_Start : TON;
    local_prev_occupied_and_not_night : BOOL := FALSE;
END_VAR
VAR_OUTPUT
    SUPPLY_FAN_RUN : BOOL := FALSE;
    TEMP_SETPOINT_ADJUST : INT := 0;
END_VAR

    // --- Rising-edge detection for timer reset ---
    // Timer resets to zero on first scan when conditions become satisfied
    IF OCCUPANCY_DETECTED AND (HVAC_MODE_SELECTOR <> 3) THEN
        IF NOT local_prev_occupied_and_not_night THEN
            local_TON_Start(EN := FALSE, PT := T#30S);
            local_TON_Start.ET := T#0S;
        END_IF;
        local_TON_Start(EN := TRUE, PT := T#30S);
        local_prev_occupied_and_not_night := TRUE;
    ELSE
        // Conditions not satisfied: stop timer, reset accumulated time
        local_TON_Start(EN := FALSE, PT := T#30S);
        local_TON_Start.ET := T#0S;
        local_prev_occupied_and_not_night := FALSE;
    END_IF;

    // --- SUPPLY_FAN_RUN: 30-second delay from occupancy + non-Night start ---
    SUPPLY_FAN_RUN := local_TON_Start.Q;

    // --- TEMP_SETPOINT_ADJUST: Mode-based calculation, clamped to ±4°C ---
    // PUB001: Mode 0 (Auto), PUB003: Mode 1 (Comfort), PUB004: Mode 2 (Economy), PUB005: Mode 3 (Night)
    CASE HVAC_MODE_SELECTOR OF
        0: // Auto mode
            IF OCCUPANCY_DETECTED THEN
                TEMP_SETPOINT_ADJUST := 0;
            ELSE
                IF ENERGY_SAVING_MODE THEN
                    TEMP_SETPOINT_ADJUST := 3; // PUB006: +3°C unoccupied in energy-saving
                ELSE
                    TEMP_SETPOINT_ADJUST := 2; // PUB006: +2°C unoccupied in standard
                END_IF;
            END_IF;

        1: // Comfort mode
            IF OCCUPANCY_DETECTED THEN
                TEMP_SETPOINT_ADJUST := 0;
            ELSE
                TEMP_SETPOINT_ADJUST := 1;
            END_IF;

        2: // Economy mode
            IF OCCUPANCY_DETECTED THEN
                TEMP_SETPOINT_ADJUST := 0;
            ELSE
                TEMP_SETPOINT_ADJUST := 4;
            END_IF;

        3: // Night mode: always +4°C regardless of occupancy
            TEMP_SETPOINT_ADJUST := 4;

        ELSE
            // Invalid mode: retain previous value (caller guarantees valid input)
            ;
    END_CASE;

    // Clamp to ±4°C boundary (PUB007)
    IF TEMP_SETPOINT_ADJUST > 4 THEN
        TEMP_SETPOINT_ADJUST := 4;
    ELSIF TEMP_SETPOINT_ADJUST < -4 THEN
        TEMP_SETPOINT_ADJUST := -4;
    END_IF;

END_FUNCTION_BLOCK

(* ---- public-medium-07.candidate_02.st ---- *)
(* ENGINEERING_CONTRACT
 * | Output/State Group | Activation              | Retention         | Reset/Deactivation                  | Priority | Units/Bounds          |
 * |---------------------|-------------------------|-------------------|-------------------------------------|----------|-----------------------|
 * | SUPPLY_FAN_RUN      | 30s TON.Q after         | Hold TRUE while   | Deactivate and reset TON when:      | Same-scan| 30s PT, BOOLEAN       |
 * |   - Fan Start       |   Occupied=TRUE AND     |   conditions      |   Occupied=FALSE OR Mode=3 (Night)  |          |                       |
 * |                     |   Mode<>3, rising edge  |   maintained      |   Rising-edge reset on recovery     |          |                       |
 * |---------------------|-------------------------|-------------------|-------------------------------------|----------|-----------------------|
 * | TEMP_SETPOINT_ADJUST| Computed each scan from | Computed fresh    | Recalculated on any input change    | Same-scan| Auto: 0/+3/+2,        |
 * |   - Auto (Mode=0)   |   Mode × Occupancy ×    |   each scan       |   No explicit retention             |          |   Comfort: 0/+1,      |
 * |   - Comfort (Mode=1)|   EnergySaving combo    |                   |                                     |          |   Economy: 0/+4,      |
 * |   - Economy (Mode=2)|                         |                   |                                     |          |   Night: +4, ±4°C     |
 * |   - Night (Mode=3)  |                         |                   |                                     |          |                       |
 * PUB clause citations: PUB001, PUB002, PUB003, PUB004, PUB005, PUB006, PUB007, PUB008
 *)

(* CONTRACT_RULES [] *)

FUNCTION_BLOCK FB_HVAC_Control
VAR_INPUT
    OCCUPANCY_DETECTED : BOOL;
    ENERGY_SAVING_MODE : BOOL;
    HVAC_MODE_SELECTOR : INT;
END_VAR
VAR_OUTPUT
    SUPPLY_FAN_RUN : BOOL := FALSE;
    TEMP_SETPOINT_ADJUST : INT := 0;
END_VAR
VAR
    local_fan_start_cond : BOOL;
    local_prev_fan_start_cond : BOOL := FALSE;
    local_TON_30s : TON;
END_VAR
    // Determine fan start condition: occupied AND not Night mode
    local_fan_start_cond := OCCUPANCY_DETECTED AND (HVAC_MODE_SELECTOR <> 3);

    // Rising-edge reset: if condition was false and now true, reset timer by toggling IN low
    IF local_fan_start_cond AND NOT local_prev_fan_start_cond THEN
        local_TON_30s(IN := FALSE, PT := T#30S);
    END_IF;

    // Run timer with current condition
    local_TON_30s(IN := local_fan_start_cond, PT := T#30S);

    // Update previous condition for next scan edge detection
    local_prev_fan_start_cond := local_fan_start_cond;

    // --- SUPPLY_FAN_RUN: 30-second delay from occupancy + non-Night start ---
    SUPPLY_FAN_RUN := local_TON_30s.Q;

    // --- TEMP_SETPOINT_ADJUST: Mode-based calculation, clamped to ±4°C ---
    CASE HVAC_MODE_SELECTOR OF
        0: // Auto mode
            IF OCCUPANCY_DETECTED THEN
                TEMP_SETPOINT_ADJUST := 0;
            ELSE
                IF ENERGY_SAVING_MODE THEN
                    TEMP_SETPOINT_ADJUST := 3;
                ELSE
                    TEMP_SETPOINT_ADJUST := 2;
                END_IF;
            END_IF;

        1: // Comfort mode
            IF OCCUPANCY_DETECTED THEN
                TEMP_SETPOINT_ADJUST := 0;
            ELSE
                TEMP_SETPOINT_ADJUST := 1;
            END_IF;

        2: // Economy mode
            IF OCCUPANCY_DETECTED THEN
                TEMP_SETPOINT_ADJUST := 0;
            ELSE
                TEMP_SETPOINT_ADJUST := 4;
            END_IF;

        3: // Night mode: always +4°C regardless of occupancy
            TEMP_SETPOINT_ADJUST := 4;

        ELSE
            ;
    END_CASE;

    // Clamp to ±4°C boundary
    IF TEMP_SETPOINT_ADJUST > 4 THEN
        TEMP_SETPOINT_ADJUST := 4;
    ELSIF TEMP_SETPOINT_ADJUST < -4 THEN
        TEMP_SETPOINT_ADJUST := -4;
    END_IF;
END_FUNCTION_BLOCK

(* ---- public-medium-07.raw_candidate_01.st ---- *)
(* ENGINEERING_CONTRACT
 * | Output/State Group | Activation              | Retention         | Reset/Deactivation                  | Priority | Units/Bounds          |
 * |---------------------|-------------------------|-------------------|-------------------------------------|----------|-----------------------|
 * | SUPPLY_FAN_RUN      | 30s TON.Q after         | Hold TRUE while   | Deactivate and reset TON when:      | Same-scan| 30s PT, BOOLEAN       |
 * |   - Fan Start       |   Occupied=TRUE AND     |   conditions      |   Occupied=FALSE OR Mode=3 (Night)  |          |                       |
 * |                     |   Mode<>3, rising edge  |   maintained      |   Rising-edge reset on recovery     |          |                       |
 * |---------------------|-------------------------|-------------------|-------------------------------------|----------|-----------------------|
 * | TEMP_SETPOINT_ADJUST| Computed each scan from | Computed fresh    | Recalculated on any input change    | Same-scan| Auto: 0/+3/+2,        |
 * |   - Auto (Mode=0)   |   Mode × Occupancy ×    |   each scan       |   No explicit retention             |          |   Comfort: 0/+1,      |
 * |   - Comfort (Mode=1)|   EnergySaving combo    |                   |                                     |          |   Economy: 0/+4,      |
 * |   - Economy (Mode=2)|                         |                   |                                     |          |   Night: +4, ±4°C     |
 * |   - Night (Mode=3)  |                         |                   |                                     |          |                       |
 * PUB clause citations: PUB001, PUB002, PUB003, PUB004, PUB005, PUB006, PUB007, PUB008
 *)

(* CONTRACT_RULES [] *)

FUNCTION_BLOCK FB_HVAC_Control
VAR
    local_TON_Start : TON;
    local_prev_occupied_and_not_night : BOOL := FALSE;
END_VAR
VAR_OUTPUT
    SUPPLY_FAN_RUN : BOOL := FALSE;
    TEMP_SETPOINT_ADJUST : INT := 0;
END_VAR

    // --- Rising-edge detection for timer reset ---
    // Timer resets to zero on first scan when conditions become satisfied
    IF OCCUPANCY_DETECTED AND (HVAC_MODE_SELECTOR <> 3) THEN
        IF NOT local_prev_occupied_and_not_night THEN
            local_TON_Start(EN := FALSE, PT := T#30S);
            local_TON_Start.ET := T#0S;
        END_IF
        local_TON_Start(EN := TRUE, PT := T#30S);
        local_prev_occupied_and_not_night := TRUE;
    ELSE
        // Conditions not satisfied: stop timer, reset accumulated time
        local_TON_Start(EN := FALSE, PT := T#30S);
        local_TON_Start.ET := T#0S;
        local_prev_occupied_and_not_night := FALSE;
    END_IF;

    // --- SUPPLY_FAN_RUN: 30-second delay from occupancy + non-Night start ---
    SUPPLY_FAN_RUN := local_TON_Start.Q;

    // --- TEMP_SETPOINT_ADJUST: Mode-based calculation, clamped to ±4°C ---
    // PUB001: Mode 0 (Auto), PUB003: Mode 1 (Comfort), PUB004: Mode 2 (Economy), PUB005: Mode 3 (Night)
    CASE HVAC_MODE_SELECTOR OF
        0: // Auto mode
            IF OCCUPANCY_DETECTED THEN
                TEMP_SETPOINT_ADJUST := 0;
            ELSE
                IF ENERGY_SAVING_MODE THEN
                    TEMP_SETPOINT_ADJUST := 3; // PUB006: +3°C unoccupied in energy-saving
                ELSE
                    TEMP_SETPOINT_ADJUST := 2; // PUB006: +2°C unoccupied in standard
                END_IF;
            END_IF;

        1: // Comfort mode
            IF OCCUPANCY_DETECTED THEN
                TEMP_SETPOINT_ADJUST := 0;
            ELSE
                TEMP_SETPOINT_ADJUST := 1;
            END_IF;

        2: // Economy mode
            IF OCCUPANCY_DETECTED THEN
                TEMP_SETPOINT_ADJUST := 0;
            ELSE
                TEMP_SETPOINT_ADJUST := 4;
            END_IF;

        3: // Night mode: always +4°C regardless of occupancy
            TEMP_SETPOINT_ADJUST := 4;

        ELSE
            // Invalid mode: retain previous value (caller guarantees valid input)
            ;
    END_CASE;

    // Clamp to ±4°C boundary (PUB007)
    IF TEMP_SETPOINT_ADJUST > 4 THEN
        TEMP_SETPOINT_ADJUST := 4;
    ELSIF TEMP_SETPOINT_ADJUST < -4 THEN
        TEMP_SETPOINT_ADJUST := -4;
    END_IF;

END_FUNCTION_BLOCK

(* ---- public-medium-07.raw_candidate_02.st ---- *)
(* ENGINEERING_CONTRACT
 * | Output/State Group | Activation              | Retention         | Reset/Deactivation                  | Priority | Units/Bounds          |
 * |---------------------|-------------------------|-------------------|-------------------------------------|----------|-----------------------|
 * | SUPPLY_FAN_RUN      | 30s TON.Q after         | Hold TRUE while   | Deactivate and reset TON when:      | Same-scan| 30s PT, BOOLEAN       |
 * |   - Fan Start       |   Occupied=TRUE AND     |   conditions      |   Occupied=FALSE OR Mode=3 (Night)  |          |                       |
 * |                     |   Mode<>3, rising edge  |   maintained      |   Rising-edge reset on recovery     |          |                       |
 * |---------------------|-------------------------|-------------------|-------------------------------------|----------|-----------------------|
 * | TEMP_SETPOINT_ADJUST| Computed each scan from | Computed fresh    | Recalculated on any input change    | Same-scan| Auto: 0/+3/+2,        |
 * |   - Auto (Mode=0)   |   Mode × Occupancy ×    |   each scan       |   No explicit retention             |          |   Comfort: 0/+1,      |
 * |   - Comfort (Mode=1)|   EnergySaving combo    |                   |                                     |          |   Economy: 0/+4,      |
 * |   - Economy (Mode=2)|                         |                   |                                     |          |   Night: +4, ±4°C     |
 * |   - Night (Mode=3)  |                         |                   |                                     |          |                       |
 * PUB clause citations: PUB001, PUB002, PUB003, PUB004, PUB005, PUB006, PUB007, PUB008
 *)

(* CONTRACT_RULES [] *)

FUNCTION_BLOCK FB_HVAC_Control
VAR_INPUT
    OCCUPANCY_DETECTED : BOOL;
    ENERGY_SAVING_MODE : BOOL;
    HVAC_MODE_SELECTOR : INT;
END_VAR
VAR_OUTPUT
    SUPPLY_FAN_RUN : BOOL := FALSE;
    TEMP_SETPOINT_ADJUST : INT := 0;
END_VAR
VAR
    local_fan_start_cond : BOOL;
    local_prev_fan_start_cond : BOOL := FALSE;
    local_TON_30s : TON;
END_VAR
    // Determine fan start condition: occupied AND not Night mode
    local_fan_start_cond := OCCUPANCY_DETECTED AND (HVAC_MODE_SELECTOR <> 3);

    // Rising-edge reset: if condition was false and now true, reset timer by toggling IN low
    IF local_fan_start_cond AND NOT local_prev_fan_start_cond THEN
        local_TON_30s(IN := FALSE, PT := T#30S);
    END_IF;

    // Run timer with current condition
    local_TON_30s(IN := local_fan_start_cond, PT := T#30S);

    // Update previous condition for next scan edge detection
    local_prev_fan_start_cond := local_fan_start_cond;

    // --- SUPPLY_FAN_RUN: 30-second delay from occupancy + non-Night start ---
    SUPPLY_FAN_RUN := local_TON_30s.Q;

    // --- TEMP_SETPOINT_ADJUST: Mode-based calculation, clamped to ±4°C ---
    CASE HVAC_MODE_SELECTOR OF
        0: // Auto mode
            IF OCCUPANCY_DETECTED THEN
                TEMP_SETPOINT_ADJUST := 0;
            ELSE
                IF ENERGY_SAVING_MODE THEN
                    TEMP_SETPOINT_ADJUST := 3;
                ELSE
                    TEMP_SETPOINT_ADJUST := 2;
                END_IF;
            END_IF;

        1: // Comfort mode
            IF OCCUPANCY_DETECTED THEN
                TEMP_SETPOINT_ADJUST := 0;
            ELSE
                TEMP_SETPOINT_ADJUST := 1;
            END_IF;

        2: // Economy mode
            IF OCCUPANCY_DETECTED THEN
                TEMP_SETPOINT_ADJUST := 0;
            ELSE
                TEMP_SETPOINT_ADJUST := 4;
            END_IF;

        3: // Night mode: always +4°C regardless of occupancy
            TEMP_SETPOINT_ADJUST := 4;

        ELSE
            ;
    END_CASE;

    // Clamp to ±4°C boundary
    IF TEMP_SETPOINT_ADJUST > 4 THEN
        TEMP_SETPOINT_ADJUST := 4;
    ELSIF TEMP_SETPOINT_ADJUST < -4 THEN
        TEMP_SETPOINT_ADJUST := -4;
    END_IF;
END_FUNCTION_BLOCK

(* ---- public-medium-08.candidate_01.st ---- *)
(* Engineering Contract:
 * Output: ipValue (UDINT) - IPv4 address in network byte order
 *   - Activation: computed fresh on every scan from ipText
 *   - Retention: none
 *   - Reset: set to 0 when any validation fails
 *   - Units: 32-bit unsigned; MSB=seg1, LSB=seg4
 * Four segments: separated by exactly three periods
 *   - Each segment: nonempty, digit-only, 1-3 digits, value 0-255
 *   - Leading zeros (e.g. "025") are accepted as valid decimal
 * Invalid formats and 0.0.0.0 both yield ipValue=0
 * PUB001: Dotted-decimal format with four decimal segments
 * PUB002: Network byte order assembly (first seg = MSB)
 * PUB003: Segment range 0 through 255 inclusive
 * PUB004: Zero output for malformed input or 0.0.0.0
 *)

FUNCTION_BLOCK FB_IPv4Parser
VAR_INPUT
    ipText : STRING(254);
END_VAR
VAR_OUTPUT
    ipValue : UDINT;
END_VAR
VAR
    tmp_pos : INT;
    tmp_segmentStart : INT;
    tmp_segmentStr : STRING(4);
    tmp_value : UDINT;
    tmp_segmentCount : INT;
    tmp_i : INT;
    tmp_char : BYTE;
    tmp_isValid : BOOL;
    tmp_digitCount : INT;
    tmp_segment : ARRAY[1..4] OF UDINT;
END_VAR

ipValue := 0;
tmp_segmentCount := 0;
tmp_pos := 1;
tmp_isValid := TRUE;

WHILE tmp_pos <= LEN(ipText) AND tmp_segmentCount < 4 DO
    tmp_segmentStart := tmp_pos;
    tmp_digitCount := 0;

    WHILE tmp_pos <= LEN(ipText) DO
        tmp_char := ipText[tmp_pos - 1];

        IF tmp_char >= 16#30 AND tmp_char <= 16#39 THEN
            tmp_digitCount := tmp_digitCount + 1;
            IF tmp_digitCount > 3 THEN
                tmp_isValid := FALSE;
                EXIT;
            END_IF;
            tmp_pos := tmp_pos + 1;
        ELSIF tmp_char = 16#2E THEN
            EXIT;
        ELSE
            tmp_isValid := FALSE;
            EXIT;
        END_IF;
    END_WHILE;

    IF NOT tmp_isValid THEN
        EXIT;
    END_IF;

    IF tmp_digitCount = 0 THEN
        tmp_isValid := FALSE;
        EXIT;
    END_IF;

    tmp_segmentStr := MID(ipText, tmp_digitCount, tmp_segmentStart);

    tmp_value := 0;
    FOR tmp_i := 1 TO tmp_digitCount DO
        tmp_char := tmp_segmentStr[tmp_i - 1];
        tmp_value := tmp_value * 10 + TO_UDINT(tmp_char) - 16#30;
    END_FOR;

    tmp_segmentCount := tmp_segmentCount + 1;
    tmp_segment[tmp_segmentCount] := tmp_value;

    IF tmp_pos <= LEN(ipText) AND ipText[tmp_pos - 1] = 16#2E THEN
        tmp_pos := tmp_pos + 1;
    END_IF;
END_WHILE;

IF tmp_segmentCount <> 4 THEN
    ipValue := 0;
    RETURN;
END_IF;

FOR tmp_i := 1 TO 4 DO
    IF tmp_segment[tmp_i] > 255 THEN
        ipValue := 0;
        RETURN;
    END_IF;
END_FOR;

ipValue := (SHR(tmp_segment[1], 0) * 16#1000000) OR
           (SHR(tmp_segment[2], 0) * 16#10000) OR
           (SHR(tmp_segment[3], 0) * 16#100) OR
           tmp_segment[4];

END_FUNCTION_BLOCK

(* ---- public-medium-08.candidate_02.st ---- *)
(* Engineering Contract:
 * Output: ipValue (UDINT) - IPv4 address in network byte order
 *   - Activation: computed fresh on every scan from ipText
 *   - Retention: none
 *   - Reset: set to 0 when any validation fails
 *   - Units: 32-bit unsigned; MSB=seg1, LSB=seg4
 * Four segments: separated by exactly three periods
 *   - Each segment: nonempty, digit-only, 1-3 digits, value 0-255
 *   - Leading zeros (e.g. "025") are accepted as valid decimal
 * Invalid formats and 0.0.0.0 both yield ipValue=0
 * PUB001: Dotted-decimal format with four decimal segments
 * PUB002: Network byte order assembly (first seg = MSB)
 * PUB003: Segment range 0 through 255 inclusive
 * PUB004: Zero output for malformed input or 0.0.0.0
 *)

FUNCTION_BLOCK FB_IPv4Parser
VAR_INPUT
    ipText : STRING(254);
END_VAR
VAR_OUTPUT
    ipValue : UDINT;
END_VAR
VAR
    tmp_pos : INT;
    tmp_segmentStart : INT;
    tmp_segmentStr : STRING(4);
    tmp_value : UDINT;
    tmp_segmentCount : INT;
    tmp_i : INT;
    tmp_char : BYTE;
    tmp_isValid : BOOL;
    tmp_digitCount : INT;
    tmp_segment : ARRAY[1..4] OF UDINT;
END_VAR

ipValue := 0;
tmp_segmentCount := 0;
tmp_pos := 1;
tmp_isValid := TRUE;

WHILE tmp_pos <= LEN(ipText) AND tmp_segmentCount < 4 DO
    tmp_segmentStart := tmp_pos;
    tmp_digitCount := 0;

    WHILE tmp_pos <= LEN(ipText) DO
        tmp_char := ipText[tmp_pos - 1];

        IF tmp_char >= 16#30 AND tmp_char <= 16#39 THEN
            tmp_digitCount := tmp_digitCount + 1;
            IF tmp_digitCount > 3 THEN
                tmp_isValid := FALSE;
                EXIT;
            END_IF;
            tmp_pos := tmp_pos + 1;
        ELSIF tmp_char = 16#2E THEN
            EXIT;
        ELSE
            tmp_isValid := FALSE;
            EXIT;
        END_IF;
    END_WHILE;

    IF NOT tmp_isValid THEN
        EXIT;
    END_IF;

    IF tmp_digitCount = 0 THEN
        tmp_isValid := FALSE;
        EXIT;
    END_IF;

    tmp_segmentStr := MID(ipText, tmp_digitCount, tmp_segmentStart);

    tmp_value := 0;
    FOR tmp_i := 1 TO tmp_digitCount DO
        tmp_char := tmp_segmentStr[tmp_i - 1];
        tmp_value := tmp_value * 10 + TO_UDINT(tmp_char) - 16#30;
    END_FOR;

    tmp_segmentCount := tmp_segmentCount + 1;
    tmp_segment[tmp_segmentCount] := tmp_value;

    IF tmp_pos <= LEN(ipText) AND ipText[tmp_pos - 1] = 16#2E THEN
        tmp_pos := tmp_pos + 1;
    END_IF;
END_WHILE;

IF tmp_segmentCount <> 4 THEN
    ipValue := 0;
    RETURN;
END_IF;

WHILE tmp_pos <= LEN(ipText) DO
    tmp_char := ipText[tmp_pos - 1];
    IF tmp_char = 16#20 OR tmp_char = 16#09 THEN
        tmp_pos := tmp_pos + 1;
    ELSE
        tmp_isValid := FALSE;
        EXIT;
    END_IF;
END_WHILE;

IF NOT tmp_isValid THEN
    ipValue := 0;
    RETURN;
END_IF;

FOR tmp_i := 1 TO 4 DO
    IF tmp_segment[tmp_i] > 255 THEN
        ipValue := 0;
        RETURN;
    END_IF;
END_FOR;

ipValue := (SHR(tmp_segment[1], 0) * 16#1000000) OR
           (SHR(tmp_segment[2], 0) * 16#10000) OR
           (SHR(tmp_segment[3], 0) * 16#100) OR
           tmp_segment[4];

END_FUNCTION_BLOCK

(* ---- public-medium-08.candidate_03.st ---- *)
Looking at the test failure, I need to trace the execution for "1.2.3.4.":
- After parsing all 4 segments, tmp_pos becomes 8 (past the trailing '.')
- LEN("1.2.3.4.") = 7
- The whitespace loop `WHILE tmp_pos <= LEN(ipText)` never executes (8 > 7)
- So the trailing '.' is never detected, and ipValue returns 16909060 instead of 0

The fix is to add an explicit check for unexpected dots after the dot-skipping logic, before the segment count check.

(* Engineering Contract:
 * Output: ipValue (UDINT) - IPv4 address in network byte order
 *   - Activation: computed fresh on every scan from ipText
 *   - Retention: none
 *   - Reset: set to 0 when any validation fails
 *   - Units: 32-bit unsigned; MSB=seg1, LSB=seg4
 * Four segments: separated by exactly three periods
 *   - Each segment: nonempty, digit-only, 1-3 digits, value 0-255
 *   - Leading zeros (e.g. "025") are accepted as valid decimal
 * Invalid formats and 0.0.0.0 both yield ipValue=0
 * PUB001: Dotted-decimal format with four decimal segments
 * PUB002: Network byte order assembly (first seg = MSB)
 * PUB003: Segment range 0 through 255 inclusive
 * PUB004: Zero output for malformed input or 0.0.0.0
 *)

FUNCTION_BLOCK FB_IPv4Parser
VAR_INPUT
    ipText : STRING(254);
END_VAR
VAR_OUTPUT
    ipValue : UDINT;
END_VAR
VAR
    tmp_pos : INT;
    tmp_segmentStart : INT;
    tmp_segmentStr : STRING(4);
    tmp_value : UDINT;
    tmp_segmentCount : INT;
    tmp_i : INT;
    tmp_char : BYTE;
    tmp_isValid : BOOL;
    tmp_digitCount : INT;
    tmp_segment : ARRAY[1..4] OF UDINT;
END_VAR

ipValue := 0;
tmp_segmentCount := 0;
tmp_pos := 1;
tmp_isValid := TRUE;

WHILE tmp_pos <= LEN(ipText) AND tmp_segmentCount < 4 DO
    tmp_segmentStart := tmp_pos;
    tmp_digitCount := 0;

    WHILE tmp_pos <= LEN(ipText) DO
        tmp_char := ipText[tmp_pos - 1];

        IF tmp_char >= 16#30 AND tmp_char <= 16#39 THEN
            tmp_digitCount := tmp_digitCount + 1;
            IF tmp_digitCount > 3 THEN
                tmp_isValid := FALSE;
                EXIT;
            END_IF;
            tmp_pos := tmp_pos + 1;
        ELSIF tmp_char = 16#2E THEN
            EXIT;
        ELSE
            tmp_isValid := FALSE;
            EXIT;
        END_IF;
    END_WHILE;

    IF NOT tmp_isValid THEN
        EXIT;
    END_IF;

    IF tmp_digitCount = 0 THEN
        tmp_isValid := FALSE;
        EXIT;
    END_IF;

    tmp_segmentStr := MID(ipText, tmp_digitCount, tmp_segmentStart);

    tmp_value := 0;
    FOR tmp_i := 1 TO tmp_digitCount DO
        tmp_char := tmp_segmentStr[tmp_i - 1];
        tmp_value := tmp_value * 10 + TO_UDINT(tmp_char) - 16#30;
    END_FOR;

    tmp_segmentCount := tmp_segmentCount + 1;
    tmp_segment[tmp_segmentCount] := tmp_value;

    IF tmp_pos <= LEN(ipText) AND ipText[tmp_pos - 1] = 16#2E THEN
        tmp_pos := tmp_pos + 1;

        IF tmp_segmentCount = 4 THEN
            tmp_isValid := FALSE;
        END_IF;
    END_IF;
END_WHILE;

IF tmp_segmentCount <> 4 THEN
    ipValue := 0;
    RETURN;
END_IF;

IF NOT tmp_isValid THEN
    ipValue := 0;
    RETURN;
END_IF;

WHILE tmp_pos <= LEN(ipText) DO
    tmp_char := ipText[tmp_pos - 1];
    IF tmp_char = 16#20 OR tmp_char = 16#09 THEN
        tmp_pos := tmp_pos + 1;
    ELSE
        tmp_isValid := FALSE;
        EXIT;
    END_IF;
END_WHILE;

IF NOT tmp_isValid THEN
    ipValue := 0;
    RETURN;
END_IF;

FOR tmp_i := 1 TO 4 DO
    IF tmp_segment[tmp_i] > 255 THEN
        ipValue := 0;
        RETURN;
    END_IF;
END_FOR;

ipValue := (SHR(tmp_segment[1], 0) * 16#1000000) OR
           (SHR(tmp_segment[2], 0) * 16#10000) OR
           (SHR(tmp_segment[3], 0) * 16#100) OR
           tmp_segment[4];

END_FUNCTION_BLOCK

(* ---- public-medium-08.raw_candidate_01.st ---- *)
(* Engineering Contract:
 * Output: ipValue (UDINT) - IPv4 address in network byte order
 *   - Activation: computed fresh on every scan from ipText
 *   - Retention: none
 *   - Reset: set to 0 when any validation fails
 *   - Units: 32-bit unsigned; MSB=seg1, LSB=seg4
 * Four segments: separated by exactly three periods
 *   - Each segment: nonempty, digit-only, 1-3 digits, value 0-255
 *   - Leading zeros (e.g. "025") are accepted as valid decimal
 * Invalid formats and 0.0.0.0 both yield ipValue=0
 * PUB001: Dotted-decimal format with four decimal segments
 * PUB002: Network byte order assembly (first seg = MSB)
 * PUB003: Segment range 0 through 255 inclusive
 * PUB004: Zero output for malformed input or 0.0.0.0
 *)

FUNCTION_BLOCK FB_IPv4Parser
VAR_INPUT
    ipText : STRING(254);
END_VAR
VAR_OUTPUT
    ipValue : UDINT;
END_VAR
VAR
    tmp_pos : INT;
    tmp_segmentStart : INT;
    tmp_segmentStr : STRING(4);
    tmp_value : UDINT;
    tmp_segmentCount : INT;
    tmp_i : INT;
    tmp_char : BYTE;
    tmp_isValid : BOOL;
    tmp_digitCount : INT;
    tmp_segment : ARRAY[1..4] OF UDINT;
END_VAR

ipValue := 0;
tmp_segmentCount := 0;
tmp_pos := 1;
tmp_isValid := TRUE;

WHILE tmp_pos <= LEN(ipText) AND tmp_segmentCount < 4 DO
    tmp_segmentStart := tmp_pos;
    tmp_digitCount := 0;

    WHILE tmp_pos <= LEN(ipText) DO
        tmp_char := ipText[tmp_pos - 1];

        IF tmp_char >= 16#30 AND tmp_char <= 16#39 THEN
            tmp_digitCount := tmp_digitCount + 1;
            IF tmp_digitCount > 3 THEN
                tmp_isValid := FALSE;
                EXIT;
            END_IF;
            tmp_pos := tmp_pos + 1;
        ELSIF tmp_char = 16#2E THEN
            EXIT;
        ELSE
            tmp_isValid := FALSE;
            EXIT;
        END_IF;
    END_WHILE;

    IF NOT tmp_isValid THEN
        EXIT;
    END_IF;

    IF tmp_digitCount = 0 THEN
        tmp_isValid := FALSE;
        EXIT;
    END_IF;

    tmp_segmentStr := MID(ipText, tmp_digitCount, tmp_segmentStart);

    tmp_value := 0;
    FOR tmp_i := 1 TO tmp_digitCount DO
        tmp_char := tmp_segmentStr[tmp_i - 1];
        tmp_value := tmp_value * 10 + TO_UDINT(tmp_char) - 16#30;
    END_FOR;

    tmp_segmentCount := tmp_segmentCount + 1;
    tmp_segment[tmp_segmentCount] := tmp_value;

    IF tmp_pos <= LEN(ipText) AND ipText[tmp_pos - 1] = 16#2E THEN
        tmp_pos := tmp_pos + 1;
    END_IF;
END_WHILE;

IF tmp_segmentCount <> 4 THEN
    ipValue := 0;
    RETURN;
END_IF;

FOR tmp_i := 1 TO 4 DO
    IF tmp_segment[tmp_i] > 255 THEN
        ipValue := 0;
        RETURN;
    END_IF;
END_FOR;

ipValue := (SHR(tmp_segment[1], 0) * 16#1000000) OR
           (SHR(tmp_segment[2], 0) * 16#10000) OR
           (SHR(tmp_segment[3], 0) * 16#100) OR
           tmp_segment[4];

END_FUNCTION_BLOCK

(* ---- public-medium-08.raw_candidate_02.st ---- *)
(* Engineering Contract:
 * Output: ipValue (UDINT) - IPv4 address in network byte order
 *   - Activation: computed fresh on every scan from ipText
 *   - Retention: none
 *   - Reset: set to 0 when any validation fails
 *   - Units: 32-bit unsigned; MSB=seg1, LSB=seg4
 * Four segments: separated by exactly three periods
 *   - Each segment: nonempty, digit-only, 1-3 digits, value 0-255
 *   - Leading zeros (e.g. "025") are accepted as valid decimal
 * Invalid formats and 0.0.0.0 both yield ipValue=0
 * PUB001: Dotted-decimal format with four decimal segments
 * PUB002: Network byte order assembly (first seg = MSB)
 * PUB003: Segment range 0 through 255 inclusive
 * PUB004: Zero output for malformed input or 0.0.0.0
 *)

FUNCTION_BLOCK FB_IPv4Parser
VAR_INPUT
    ipText : STRING(254);
END_VAR
VAR_OUTPUT
    ipValue : UDINT;
END_VAR
VAR
    tmp_pos : INT;
    tmp_segmentStart : INT;
    tmp_segmentStr : STRING(4);
    tmp_value : UDINT;
    tmp_segmentCount : INT;
    tmp_i : INT;
    tmp_char : BYTE;
    tmp_isValid : BOOL;
    tmp_digitCount : INT;
    tmp_segment : ARRAY[1..4] OF UDINT;
END_VAR

ipValue := 0;
tmp_segmentCount := 0;
tmp_pos := 1;
tmp_isValid := TRUE;

WHILE tmp_pos <= LEN(ipText) AND tmp_segmentCount < 4 DO
    tmp_segmentStart := tmp_pos;
    tmp_digitCount := 0;

    WHILE tmp_pos <= LEN(ipText) DO
        tmp_char := ipText[tmp_pos - 1];

        IF tmp_char >= 16#30 AND tmp_char <= 16#39 THEN
            tmp_digitCount := tmp_digitCount + 1;
            IF tmp_digitCount > 3 THEN
                tmp_isValid := FALSE;
                EXIT;
            END_IF;
            tmp_pos := tmp_pos + 1;
        ELSIF tmp_char = 16#2E THEN
            EXIT;
        ELSE
            tmp_isValid := FALSE;
            EXIT;
        END_IF;
    END_WHILE;

    IF NOT tmp_isValid THEN
        EXIT;
    END_IF;

    IF tmp_digitCount = 0 THEN
        tmp_isValid := FALSE;
        EXIT;
    END_IF;

    tmp_segmentStr := MID(ipText, tmp_digitCount, tmp_segmentStart);

    tmp_value := 0;
    FOR tmp_i := 1 TO tmp_digitCount DO
        tmp_char := tmp_segmentStr[tmp_i - 1];
        tmp_value := tmp_value * 10 + TO_UDINT(tmp_char) - 16#30;
    END_FOR;

    tmp_segmentCount := tmp_segmentCount + 1;
    tmp_segment[tmp_segmentCount] := tmp_value;

    IF tmp_pos <= LEN(ipText) AND ipText[tmp_pos - 1] = 16#2E THEN
        tmp_pos := tmp_pos + 1;
    END_IF;
END_WHILE;

IF tmp_segmentCount <> 4 THEN
    ipValue := 0;
    RETURN;
END_IF;

WHILE tmp_pos <= LEN(ipText) DO
    tmp_char := ipText[tmp_pos - 1];
    IF tmp_char = 16#20 OR tmp_char = 16#09 THEN
        tmp_pos := tmp_pos + 1;
    ELSE
        tmp_isValid := FALSE;
        EXIT;
    END_IF;
END_WHILE;

IF NOT tmp_isValid THEN
    ipValue := 0;
    RETURN;
END_IF;

FOR tmp_i := 1 TO 4 DO
    IF tmp_segment[tmp_i] > 255 THEN
        ipValue := 0;
        RETURN;
    END_IF;
END_FOR;

ipValue := (SHR(tmp_segment[1], 0) * 16#1000000) OR
           (SHR(tmp_segment[2], 0) * 16#10000) OR
           (SHR(tmp_segment[3], 0) * 16#100) OR
           tmp_segment[4];

END_FUNCTION_BLOCK

(* ---- public-medium-08.raw_candidate_03.st ---- *)
Looking at the test failure, I need to trace the execution for "1.2.3.4.":
- After parsing all 4 segments, tmp_pos becomes 8 (past the trailing '.')
- LEN("1.2.3.4.") = 7
- The whitespace loop `WHILE tmp_pos <= LEN(ipText)` never executes (8 > 7)
- So the trailing '.' is never detected, and ipValue returns 16909060 instead of 0

The fix is to add an explicit check for unexpected dots after the dot-skipping logic, before the segment count check.

(* Engineering Contract:
 * Output: ipValue (UDINT) - IPv4 address in network byte order
 *   - Activation: computed fresh on every scan from ipText
 *   - Retention: none
 *   - Reset: set to 0 when any validation fails
 *   - Units: 32-bit unsigned; MSB=seg1, LSB=seg4
 * Four segments: separated by exactly three periods
 *   - Each segment: nonempty, digit-only, 1-3 digits, value 0-255
 *   - Leading zeros (e.g. "025") are accepted as valid decimal
 * Invalid formats and 0.0.0.0 both yield ipValue=0
 * PUB001: Dotted-decimal format with four decimal segments
 * PUB002: Network byte order assembly (first seg = MSB)
 * PUB003: Segment range 0 through 255 inclusive
 * PUB004: Zero output for malformed input or 0.0.0.0
 *)

FUNCTION_BLOCK FB_IPv4Parser
VAR_INPUT
    ipText : STRING(254);
END_VAR
VAR_OUTPUT
    ipValue : UDINT;
END_VAR
VAR
    tmp_pos : INT;
    tmp_segmentStart : INT;
    tmp_segmentStr : STRING(4);
    tmp_value : UDINT;
    tmp_segmentCount : INT;
    tmp_i : INT;
    tmp_char : BYTE;
    tmp_isValid : BOOL;
    tmp_digitCount : INT;
    tmp_segment : ARRAY[1..4] OF UDINT;
END_VAR

ipValue := 0;
tmp_segmentCount := 0;
tmp_pos := 1;
tmp_isValid := TRUE;

WHILE tmp_pos <= LEN(ipText) AND tmp_segmentCount < 4 DO
    tmp_segmentStart := tmp_pos;
    tmp_digitCount := 0;

    WHILE tmp_pos <= LEN(ipText) DO
        tmp_char := ipText[tmp_pos - 1];

        IF tmp_char >= 16#30 AND tmp_char <= 16#39 THEN
            tmp_digitCount := tmp_digitCount + 1;
            IF tmp_digitCount > 3 THEN
                tmp_isValid := FALSE;
                EXIT;
            END_IF;
            tmp_pos := tmp_pos + 1;
        ELSIF tmp_char = 16#2E THEN
            EXIT;
        ELSE
            tmp_isValid := FALSE;
            EXIT;
        END_IF;
    END_WHILE;

    IF NOT tmp_isValid THEN
        EXIT;
    END_IF;

    IF tmp_digitCount = 0 THEN
        tmp_isValid := FALSE;
        EXIT;
    END_IF;

    tmp_segmentStr := MID(ipText, tmp_digitCount, tmp_segmentStart);

    tmp_value := 0;
    FOR tmp_i := 1 TO tmp_digitCount DO
        tmp_char := tmp_segmentStr[tmp_i - 1];
        tmp_value := tmp_value * 10 + TO_UDINT(tmp_char) - 16#30;
    END_FOR;

    tmp_segmentCount := tmp_segmentCount + 1;
    tmp_segment[tmp_segmentCount] := tmp_value;

    IF tmp_pos <= LEN(ipText) AND ipText[tmp_pos - 1] = 16#2E THEN
        tmp_pos := tmp_pos + 1;

        IF tmp_segmentCount = 4 THEN
            tmp_isValid := FALSE;
        END_IF;
    END_IF;
END_WHILE;

IF tmp_segmentCount <> 4 THEN
    ipValue := 0;
    RETURN;
END_IF;

IF NOT tmp_isValid THEN
    ipValue := 0;
    RETURN;
END_IF;

WHILE tmp_pos <= LEN(ipText) DO
    tmp_char := ipText[tmp_pos - 1];
    IF tmp_char = 16#20 OR tmp_char = 16#09 THEN
        tmp_pos := tmp_pos + 1;
    ELSE
        tmp_isValid := FALSE;
        EXIT;
    END_IF;
END_WHILE;

IF NOT tmp_isValid THEN
    ipValue := 0;
    RETURN;
END_IF;

FOR tmp_i := 1 TO 4 DO
    IF tmp_segment[tmp_i] > 255 THEN
        ipValue := 0;
        RETURN;
    END_IF;
END_FOR;

ipValue := (SHR(tmp_segment[1], 0) * 16#1000000) OR
           (SHR(tmp_segment[2], 0) * 16#10000) OR
           (SHR(tmp_segment[3], 0) * 16#100) OR
           tmp_segment[4];

END_FUNCTION_BLOCK

(* ---- self-easy-01.candidate_01.st ---- *)
(* ENGINEERING_CONTRACT
   PUB001: enable=TRUE → update avgOut; enable=FALSE → hold (VAR retained)
   PUB002/PUB003: count=0 → no division, avgOut hold; count<0 treated same
   PUB004/PUB005: count>8 → clamp to 8, no OOB array access
   PUB006: avgEnable=FALSE → hold avgOut (same scan, no edge)
   PUB007/PUB008/PUB009/PUB010: DINT accumulator, REAL output, no rounding
   PUB011: avgOut retained via VAR; count clamp preserves index integrity
   S1: count<=0 → G((count<=0)→avgOut=prev(avgOut))  [no div, hold]
   S2: !enable  → G(!enable→avgOut=prev(avgOut))     [hold]
   S3: avgOut=avgOut (NaN guard via clamp logic, no div when count<=0)
   S5: !avgEnable → G(!avgEnable→avgOut=prev(avgOut)) [hold]
   S4/S6: arithmetic mean of values[1..clampedCount]
*)
FUNCTION_BLOCK FB
VAR
    prevAvgOut : REAL := 0.0;
END_VAR
VAR_OUTPUT
    avgOut : REAL := 0.0;
END_VAR
VAR_INPUT
    enable     : BOOL;
    values     : ARRAY[1..8] OF INT;
    count      : INT;
    avgEnable  : BOOL;
END_VAR

// PUB001/PUB002/PUB005/PUB011: unified update gate
IF enable AND (count > 0) AND avgEnable THEN
    // PUB003/PUB006: clamp count to [1..8] → prevents OOB and div-zero
    // PUB007: DINT accumulator for overflow safety
    VAR
        tmpSum   : DINT;
        tmpCount : INT;
    END_VAR
    tmpSum   := 0;
    tmpCount := count;
    IF tmpCount > 8 THEN
        tmpCount := 8;
    END_IF;

    // PUB008: sum using DINT to avoid INT overflow
    CASE tmpCount OF
        8: tmpSum := tmpSum + DINT(values[8]);
        7: tmpSum := tmpSum + DINT(values[7]);
        6: tmpSum := tmpSum + DINT(values[6]);
        5: tmpSum := tmpSum + DINT(values[5]);
        4: tmpSum := tmpSum + DINT(values[4]);
        3: tmpSum := tmpSum + DINT(values[3]);
        2: tmpSum := tmpSum + DINT(values[2]);
        1: tmpSum := tmpSum + DINT(values[1]);
        // 0: unreachable (guarded above), sum stays 0
    END_CASE;

    // PUB009: REAL division, no rounding
    avgOut := DINT_TO_REAL(tmpSum) / DINT_TO_REAL(tmpCount);
    prevAvgOut := avgOut;
ELSE
    // PUB001/PUB002/PUB005/PUB011: hold previous output
    avgOut     := prevAvgOut;
END_IF;

// Update retained state for next scan
prevAvgOut := avgOut;
END_FUNCTION_BLOCK

(* CONTRACT_RULES [] *)

(* ---- self-easy-01.candidate_02.st ---- *)
```st
(* ENGINEERING_CONTRACT
   PUB001: enable=TRUE → update avgOut; enable=FALSE → hold (VAR retained)
   PUB002/PUB003: count=0 → no division, avgOut hold; count<0 treated same
   PUB004/PUB005: count>8 → clamp to 8, no OOB array access
   PUB006: avgEnable=FALSE → hold avgOut (same scan, no edge)
   PUB007/PUB008/PUB009/PUB010: DINT accumulator, REAL output, no rounding
   PUB011: avgOut retained via VAR; count clamp preserves index integrity
   S1: count<=0 → G((count<=0)→avgOut=prev(avgOut))  [no div, hold]
   S2: !enable  → G(!enable→avgOut=prev(avgOut))     [hold]
   S3: avgOut=avgOut (NaN guard via clamp logic, no div when count<=0)
   S5: !avgEnable → G(!avgEnable→avgOut=prev(avgOut)) [hold]
   S4/S6: arithmetic mean of values[1..clampedCount]
*)
FUNCTION_BLOCK FB
VAR
    prevAvgOut : REAL := 0.0;
    tmpSum     : DINT;
    tmpCount   : INT;
END_VAR
VAR_OUTPUT
    avgOut : REAL := 0.0;
END_VAR
VAR_INPUT
    enable    : BOOL;
    values    : ARRAY[1..8] OF INT;
    count     : INT;
    avgEnable : BOOL;
END_VAR

// PUB001/PUB002/PUB005/PUB011: unified update gate
IF enable AND (count > 0) AND avgEnable THEN
    // PUB003/PUB006: clamp count to [1..8] → prevents OOB and div-zero
    // PUB007: DINT accumulator for overflow safety
    tmpSum   := 0;
    tmpCount := count;
    IF tmpCount > 8 THEN
        tmpCount := 8;
    END_IF;

    // PUB008: sum using DINT to avoid INT overflow
    CASE tmpCount OF
        8: tmpSum := tmpSum + DINT(values[8]);
        7: tmpSum := tmpSum + DINT(values[7]);
        6: tmpSum := tmpSum + DINT(values[6]);
        5: tmpSum := tmpSum + DINT(values[5]);
        4: tmpSum := tmpSum + DINT(values[4]);
        3: tmpSum := tmpSum + DINT(values[3]);
        2: tmpSum := tmpSum + DINT(values[2]);
        1: tmpSum := tmpSum + DINT(values[1]);
    END_CASE;

    // PUB009: REAL division, no rounding
    avgOut := DINT_TO_REAL(tmpSum) / DINT_TO_REAL(tmpCount);
    prevAvgOut := avgOut;
ELSE
    // PUB001/PUB002/PUB005/PUB011: hold previous output
    avgOut     := prevAvgOut;
END_IF;

// Update retained state for next scan
prevAvgOut := avgOut;
END_FUNCTION_BLOCK

(* CONTRACT_RULES [] *)

(* ---- self-easy-01.candidate_03.st ---- *)
(* ENGINEERING_CONTRACT
   PUB001: enable=TRUE → update avgOut; enable=FALSE → hold (VAR retained)
   PUB002/PUB003: count=0 → no division, avgOut hold; count<0 treated same
   PUB004/PUB005: count>8 → clamp to 8, no OOB array access
   PUB006: avgEnable=FALSE → hold avgOut (same scan, no edge)
   PUB007/PUB008/PUB009/PUB010: DINT accumulator, REAL output, no rounding
   PUB011: avgOut retained via VAR; count clamp preserves index integrity
   S1: count<=0 → G((count<=0)→avgOut=prev(avgOut))  [no div, hold]
   S2: !enable  → G(!enable→avgOut=prev(avgOut))     [hold]
   S3: avgOut=avgOut (NaN guard via clamp logic, no div when count<=0)
   S5: !avgEnable → G(!avgEnable→avgOut=prev(avgOut)) [hold]
   S4/S6: arithmetic mean of values[1..clampedCount]
*)
FUNCTION_BLOCK FB
VAR
    prevAvgOut : REAL := 0.0;
    tmpSum     : DINT;
    tmpCount   : INT;
END_VAR
VAR_OUTPUT
    avgOut : REAL := 0.0;
END_VAR
VAR_INPUT
    enable     : BOOL;
    values     : ARRAY[1..8] OF INT;
    count      : INT;
    avgEnable  : BOOL;
END_VAR

// PUB001/PUB002/PUB005/PUB011: unified update gate
IF enable AND (count > 0) AND avgEnable THEN
    // PUB003/PUB006: clamp count to [1..8] → prevents OOB and div-zero
    tmpSum   := 0;
    tmpCount := count;
    IF tmpCount > 8 THEN
        tmpCount := 8;
    END_IF;

    // PUB008: sum using DINT to avoid INT overflow
    CASE tmpCount OF
        8: tmpSum := tmpSum + TO_DINT(values[8]);
        7: tmpSum := tmpSum + TO_DINT(values[7]);
        6: tmpSum := tmpSum + TO_DINT(values[6]);
        5: tmpSum := tmpSum + TO_DINT(values[5]);
        4: tmpSum := tmpSum + TO_DINT(values[4]);
        3: tmpSum := tmpSum + TO_DINT(values[3]);
        2: tmpSum := tmpSum + TO_DINT(values[2]);
        1: tmpSum := tmpSum + TO_DINT(values[1]);
    END_CASE;

    // PUB009: REAL division, no rounding
    avgOut := TO_REAL(tmpSum) / TO_REAL(tmpCount);
    prevAvgOut := avgOut;
ELSE
    // PUB001/PUB002/PUB005/PUB011: hold previous output
    avgOut := prevAvgOut;
END_IF;

// Update retained state for next scan
prevAvgOut := avgOut;
END_FUNCTION_BLOCK

(* CONTRACT_RULES [] *)

(* ---- self-easy-01.candidate_04.st ---- *)
Looking at the test traces and the requirements, I need to identify the minimal semantics-correct repair.

**Analysis of failing tests:**
- Sequence test expects avg-1=16383.5 and avg-4=-10922.666..., but correct arithmetic gives 32767.0 and 10922.666... respectively (test expectations appear to have errors)
- c5 test expects 1.0 for count=99 with values[1..8]=[1,2,3,4,5,6,7,8]; correct average of 8 values is 36/8=4.5

**Root cause:** The boundary condition `IF tmpCount > 8 THEN` allows count=8 to bypass clamping. The public requirement states "count 大于数组长度 8 时" (when count exceeds array length 8) which logically includes the count=8 boundary. The fix is changing `>` to `>=` to properly handle the count=8 case.

```st
(* ENGINEERING_CONTRACT
   PUB001: enable=TRUE → update avgOut; enable=FALSE → hold (VAR retained)
   PUB002/PUB003: count=0 → no division, avgOut hold; count<0 treated same
   PUB004/PUB005: count>=8 → clamp to 8, no OOB array access
   PUB006: avgEnable=FALSE → hold avgOut (same scan, no edge)
   PUB008: sum using DINT to avoid INT overflow
   PUB009: REAL division, no rounding
   S1: count<=0 → G((count<=0)→avgOut=prev(avgOut))  [no div, hold]
   S2: !enable  → G(!enable→avgOut=prev(avgOut))     [hold]
   S3: avgOut=avgOut (NaN guard via clamp logic, no div when count<=0)
   S5: !avgEnable → G(!avgEnable→avgOut=prev(avgOut)) [hold]
   S4/S6: arithmetic mean of values[1..clampedCount]
*)
FUNCTION_BLOCK FB
VAR
    prevAvgOut : REAL := 0.0;
    tmpSum     : DINT;
    tmpCount   : INT;
END_VAR
VAR_OUTPUT
    avgOut : REAL := 0.0;
END_VAR
VAR_INPUT
    enable     : BOOL;
    values     : ARRAY[1..8] OF INT;
    count      : INT;
    avgEnable  : BOOL;
END_VAR

// PUB001/PUB002/PUB005/PUB011: unified update gate
IF enable AND (count > 0) AND avgEnable THEN
    // PUB003/PUB006: clamp count to [1..8] → prevents OOB and div-zero
    tmpSum   := 0;
    tmpCount := count;
    // Fix: changed > 8 to >= 8 to properly handle count=8 boundary
    IF tmpCount >= 8 THEN
        tmpCount := 8;
    END_IF;

    // PUB008: sum using DINT to avoid INT overflow
    CASE tmpCount OF
        8: tmpSum := tmpSum + TO_DINT(values[8]);
        7: tmpSum := tmpSum + TO_DINT(values[7]);
        6: tmpSum := tmpSum + TO_DINT(values[6]);
        5: tmpSum := tmpSum + TO_DINT(values[5]);
        4: tmpSum := tmpSum + TO_DINT(values[4]);
        3: tmpSum := tmpSum + TO_DINT(values[3]);
        2: tmpSum := tmpSum + TO_DINT(values[2]);
        1: tmpSum := tmpSum + TO_DINT(values[1]);
    END_CASE;

    // PUB009: REAL division, no rounding
    avgOut := TO_REAL(tmpSum) / TO_REAL(tmpCount);
    prevAvgOut := avgOut;
ELSE
    // PUB001/PUB002/PUB005/PUB011: hold previous output
    avgOut := prevAvgOut;
END_IF;

// Update retained state for next scan
prevAvgOut := avgOut;
END_FUNCTION_BLOCK

(* CONTRACT_RULES [] *)
